(* IEC 61131-3 sources: test/Class/LseEasy, 1 file *)

(* ---- LseEasy.st ---- *)
#include "..\..\Source\Common\hmi_nuc.h"

(*!
<Class
	Name               = "LseEasy"
	Revision           = "1.32"
	RealtimeTask       = "false"
	CyclicTask         = "false"
	BackgroundTask     = "true"
	DefBackground      = "always"
	Sigmatek           = "true"
	OSInterface        = "false"
	HighPriority       = "false"
	Automatic          = "false"
	UpdateMode         = "Prescan"
	SharedCommandTable = "true"
	Objectsize         = "(474,120)"
	Comment            = "Class is used to operate LSE-Easy Visualization&#13;&#10;LSE-CompilerVersion: 60">
	<Channels>
		<Server Name="AccessLevel" Visualized="true" Initialize="false" WriteProtected="false" Retentive="false" Comment="server is used to disable/enable access to several inputs and buttons&#13;&#10;virtual method HmiAccess() is responsible for algorithm."/>
		<Server Name="ActHumidity" Visualized="true" Initialize="false" WriteProtected="true" Retentive="false" Comment="actual humidity"/>
		<Server Name="ActLanguage" Visualized="true" Initialize="true" DefValue="0" WriteProtected="false" Retentive="SRam" Comment="Server is used to select language&#13;&#10;use index or accurate language designator to switch over"/>
		<Server Name="ActScreen" Visualized="true" Initialize="false" WriteProtected="false" Retentive="false" Comment="server is used to show number of actual screen on hmi&#13;&#10;call write-method with accurate screennumber given by lse to force hmi to view new screen&#13;&#10;call writemethode with -2 to get screenshot from hmi (C:\hmi35.bmp)"/>
		<Server Name="ActTemperature" Visualized="true" Initialize="false" WriteProtected="true" Retentive="false" Comment="actual temperature"/>
		<Server Name="BacklightDim" Visualized="true" Initialize="false" WriteProtected="false" Retentive="false" Comment="server is used to dim backlight of hmi&#13;&#10;call writemethode with any value from 0 to 100 to dim backlight&#13;&#10;0 .... next to dark&#13;&#10;100 .. bright"/>
		<Server Name="BacklightOnOff" Visualized="false" Initialize="false" WriteProtected="false" Retentive="false" Comment="server is used to turn on/off backlight of hmi&#13;&#10;call writemethode with 0 to turn off backlight&#13;&#10;on the oter hand call writemethode with 1 to turn on backlight"/>
		<Server Name="ClassSvr" Visualized="false" Initialize="false" WriteProtected="true" Retentive="false"/>
		<Server Name="ErrorSvr" Visualized="true" Initialize="false" WriteProtected="true" Retentive="false"/>
		<Server Name="HmiHwVersion" Visualized="true" Initialize="false" WriteProtected="true" Retentive="false" Comment="is used to view hardwareversion of hmi"/>
		<Server Name="HmiOnline" Visualized="true" Initialize="false" WriteProtected="true" Retentive="false" Comment="0 ... hmi is offline&#13;&#10;1 ... hmi is online"/>
		<Server Name="HmiSwVersion" Visualized="true" Initialize="false" WriteProtected="true" Retentive="false" Comment="is used to view softwareversion (firmware) of hmi"/>
		<Server Name="LastUsage" Visualized="false" Initialize="false" WriteProtected="true" Retentive="false" Comment="server is used to display timestamp (ops.tabsolute) of last usage of hmi"/>
		<Server Name="ListVal0" Visualized="true" Initialize="false" WriteProtected="false" Retentive="false" Comment="server is used to display arbitrary scrolllist on display&#13;&#10;actual selection in list will be shown on server"/>
		<Server Name="ListVal1" Visualized="true" Initialize="false" WriteProtected="false" Retentive="false"/>
		<Server Name="LseProjectRevision" Visualized="true" Initialize="false" WriteProtected="true" Retentive="false"/>
		<Server Name="PixMap" Visualized="true" Initialize="false" WriteProtected="false" Retentive="false"/>
		<Server Name="StateSvr" Visualized="true" Initialize="false" WriteProtected="false" Retentive="false" Comment="actual state of program"/>
		<Server Name="TrendVal0" Visualized="true" Initialize="false" WriteProtected="false" Retentive="false" Comment="server is used to display trend0 on hmi&#13;&#10;call writemethod with any value from 0 to 255 to add value"/>
		<Server Name="TrendVal1" Visualized="true" Initialize="false" WriteProtected="false" Retentive="false" Comment="server is used to display trend1 on hmi&#13;&#10;call writemethod with any value from 0 to 255 to add value"/>
		<Client Name="AutoFirmwareUpdate" Required="true" Internal="false" DefValue="0" Comment="Client is used to ensure automatic update of firmware and bootloader at hmi after poweron of connected plc.&#13;&#10;Set client to 1 or 2 to enable automatic update otherwirse, when client is set to 0, automatic update is disabled.&#13;&#10;NOTE: &#13;&#10;If client is set to 1, updatefiles will be deleted after update of hmi. &#13;&#10;When client is set to 2, updatefiles will NOT be deleted after automatic update. In that case user has to disconnect device otherwise update will be performed each time after poweron.&#13;&#10;User has to place updatefiles at correct device (eg.: C:\, E:\, ...}. When updatefiles should be deleted after success make sure that device and updatefiles are not writeprotected.&#13;&#10;Use virtual methods GetUpdatePath(), GetFirmwareUpdate() and GetBootLoaderUpdate() to customize device, directory and name of updatefiles."/>
		<Client Name="BackLightOff" Required="true" Internal="false" DefValue="300000" Comment="client is used to set duration till backlight will be turned off when display is not in use&#13;&#10;timebase is milliseconds&#13;&#10;0 ... backlight is always on"/>
		<Client Name="ComPort" Required="true" Internal="false" Comment="client is used to communicate with hmi&#13;&#10;eg: connect instance of class HmiComPortCan to communicate vie canbus"/>
		<Client Name="File" Required="true" Internal="true"/>
		<Client Name="HmiChkBitList" Required="true" Internal="true"/>
		<Client Name="HmiColorMap" Required="true" Internal="true"/>
		<Client Name="HmiFont35" Required="true" Internal="true"/>
		<Client Name="HmiFontList" Required="true" Internal="true"/>
		<Client Name="HmiFontShemeList" Required="true" Internal="true"/>
		<Client Name="HmiFunctionList" Required="true" Internal="true"/>
		<Client Name="HmiFunctionList35" Required="true" Internal="true"/>
		<Client Name="HmiImage35" Required="true" Internal="true"/>
		<Client Name="HmiImageList" Required="true" Internal="true"/>
		<Client Name="HmiImageShemeList" Required="true" Internal="true"/>
		<Client Name="HmiMapFile" Required="true" Internal="true"/>
		<Client Name="HmiProject35" Required="true" Internal="true"/>
		<Client Name="HmiProjectList" Required="true" Internal="true"/>
		<Client Name="HmiScreen" Required="true" Internal="true"/>
		<Client Name="HmiSetUpList" Required="true" Internal="true"/>
		<Client Name="HmiSetupList35" Required="true" Internal="true"/>
		<Client Name="HmiShemeList35" Required="true" Internal="true"/>
		<Client Name="HmiStateBit35" Required="true" Internal="true"/>
		<Client Name="HmiT9Config" Required="true" Internal="true"/>
		<Client Name="HmiTextList" Required="true" Internal="true"/>
		<Client Name="HmiTextList35" Required="true" Internal="true"/>
		<Client Name="HmiTextShemeList" Required="true" Internal="true"/>
		<Client Name="HmiUtils" Required="true" Internal="true"/>
		<Client Name="HmiVarList" Required="true" Internal="true"/>
		<Client Name="HmiVarList35" Required="true" Internal="true"/>
		<Client Name="OverloadLight" Required="true" Internal="false" DefValue="-1" Comment="client is used to ensure overload&#13;&#10;if client is set to equal or bigger 0 all occurences of &quot;XX&quot; in variablename done with LSE will be xchanged with adequateness number of client"/>
		<Client Name="ProjectPath" Required="true" Internal="false" DefValue="0" Comment="selector for different projectpath&#13;&#10;0: C:\MPC\&#13;&#10;&gt;0: C:\Easy[Value]\ (eg.: C:\Easy123\)&#13;&#10;-1: C:\[ObjextName]\ (eg.: C:\LSEEASY1\)&#13;&#10;"/>
		<Client Name="StringLib" Required="true" Internal="true"/>
		<Client Name="TempInterval" Required="true" Internal="false" DefValue="1000" Comment="client is used to define interval of retrieving act.temperature from hmi&#13;&#10;timebase is milliseconds&#13;&#10;0 ... do not update act.temperature"/>
	</Channels>
	<Dependencies>
		<Files>
			<File Path=".\Source\Common\hmi_nuc.h" Include="true"/>
			<File Path=".\Class\LseEasy\MiniSrcData.h" Include="false"/>
			<File Path=".\Class\LseEasy\Create.h" Include="false"/>
			<File Path=".\Class\LseEasy\CreateScreen.c"/>
			<File Path=".\Class\LseEasy\CreateUtils.c"/>
		</Files>
	</Dependencies>
	<RevDoku>
		<Owner Company="sigmatek" Author="kolott"/>
		<Dokumentation Revision="1.32" Date="2021-02-26" Author="kolott" Company="sigmatek" Description="Method LseEasy::ListSetup() by parameter &apos;bottom_up&apos; expanded&#13;&#10;8D-1972: Extended size of textpuffer"/>
		<Dokumentation Revision="1.31" Date="2020-04-28" Author="kolott" Company="sigmatek" Description="New method GetLseProjectName() added&#13;&#10;DEVVIS-40, sa57116: New method T9KeyboardConfig() added"/>
		<Dokumentation Revision="1.30" Date="2019-01-24" Author="kolott" Company="sigmatek" Description="Support of HZS-251-1 and HZS352-1 incl. Humidity"/>
		<Dokumentation Revision="1.29" Date="2019-01-09" Author="kolott" Company="sigmatek" Description="Virtual method HmiOverloadLight() added to ensure userspecific change of Objectname"/>
		<Dokumentation Revision="1.28" Date="2018-10-18" Author="kolott" Company="sigmatek" Description="sa42417: more than 6 different projectpath implemented in virtual method LseEasy::GetPrjPath()"/>
		<Dokumentation Revision="1.27" Date="2018-08-27" Author="kolott" Company="sigmatek" Description="Problem &quot;Out Of Memory&quot; will end in Error &quot;Can&apos;t load LSE-Project&quot;&#13;&#10;Variable Limits at Variables will work. Overwrite Method LseEasy::VariableLimitsInUse() to enable feature"/>
		<Dokumentation Revision="1.26" Date="2018-05-24" Author="kolott" Company="sigmatek" Description="sa41119, DEVSW502: Send individual StandardFonts given by LSE to HMI as well. Fonts are used in Standard Keypads"/>
		<Dokumentation Revision="1.25" Date="2018-04-18" Author="kolott" Company="sigmatek" Description="sa40364: userspecific xchange of images done by LSE.&#13;&#10;DEVSW440: Server ActTemperature is set to 16#80000010 when HMI is offline and TemperatureValue is needed"/>
		<Dokumentation Revision="1.24" Date="2018-01-17" Author="kolott" Company="sigmatek" Description="TextList done wilt LSE will be accessible by user during runtime&#13;&#10;new virtual method HmiProjectBegin(), AddVariableByName() and AddStateBitByName() added"/>
		<Dokumentation Revision="1.23" Date="2016-09-07" Author="kolott" Company="sigmatek" Description="sa35391: new method GetLseProjectNotice() and Server LseProjectRevision added&#13;&#10;sa35411: correction in entire bytesizecomputation of HMI-project-data"/>
		<Dokumentation Revision="1.22" Date="2016-07-08" Author="kolott" Company="sigmatek" Description="new Client AutoFirmwareUpdate added to enable automatic update of firmware and bootloader at hmi after poweron"/>
		<Dokumentation Revision="1.21" Date="2016-06-22" Author="kolott" Company="sigmatek" Description="Functionality to Update BootLoader in HMI added"/>
		<Dokumentation Revision="1.20" Date="2016-05-03" Author="kolott" Company="sigmatek" Description="Betterment in rounding result at method Calc().&#13;&#10;Set and resetvalue at button will work. Firmwareversion 1.35 or higher is necessary at HMI.&#13;&#10;sa26785: compilerversion 60, property preceding zero implemented&#13;&#10;Methode UpdateString35() is done virtual"/>
		<Dokumentation Revision="1.19" Date="2016-04-23" Author="kolott" Company="sigmatek" Description="sa34276: new methode Recalculate() added to ensure recalculation from binary to physical values"/>
		<Dokumentation Revision="1.18" Date="2016-03-12" Author="kolott" Company="sigmatek" Description="functionality to display pixmap (barcode, qr code,...) on hmi added. use method SendPixMap() to view data&#13;&#10;correction of server ActLanguage when actual selection doesn&apos;t fit to loaded project (sa33823)"/>
		<Dokumentation Revision="1.17" Date="2016-02-04" Author="kolott" Company="sigmatek" Description="new virtual method IsProjectUpLoadNecessary() to customize project-upload added"/>
		<Dokumentation Revision="1.16" Date="2015-11-30" Author="kolott" Company="sigmatek" Description="new Server &quot;ListVal1&quot; to ensure use of second scrolllist on HMI"/>
		<Dokumentation Revision="1.15" Date="2015-03-17" Author="kolott" Company="sigmatek" Description="method UpdateValue35() is done &quot;virtual&quot;"/>
		<Dokumentation Revision="1.14" Date="2014-11-26" Author="kolott" Company="sigmatek" Description="new method HmiVariableExtention() used to ensure userextended modifications done in firmware of hmi&#13;&#10;view Passwordcharacter at String will work"/>
		<Dokumentation Revision="1.13" Date="2014-10-15" Author="kolott" Company="sigmatek" Description="Ability to customise HmiProject added (HmiProjectCreate(), CreateAddText(), CreateAddImage(), ListSetup(), ListCmd(), ListAddItem())"/>
		<Dokumentation Revision="1.12" Date="2014-08-13" Author="kolott" Company="sigmatek" Description="Server &quot;ListVal0&quot; is added to ensure scrollist on HMI&#13;&#10;Function &quot;UserCall&quot; added&#13;&#10;Retry added at filetransfer to HMI"/>
		<Dokumentation Revision="1.11" Date="2014-08-07" Author="kolott" Company="sigmatek" Description="Server of type ENUM will work as well"/>
		<Dokumentation Revision="1.10" Date="2014-06-02" Author="kolott" Company="sigmatek" Description="Method &quot;UpdateTemperature35&quot; is virtual to ensure correction of actual HMI-Temperature&#13;&#10;Correction: Display of Unicode-String always started with character &apos;?&apos;"/>
		<Dokumentation Revision="1.9" Date="2014-04-28" Author="kolott" Company="sigmatek" Description="call of function &quot;Function Block&quot; activated&#13;&#10;view of Circle + Pie added"/>
		<Dokumentation Revision="1.8" Date="2014-04-14" Author="kolott" Company="sigmatek" Description="betterment in Offline-Mode when HMI (display) is not connected&#13;&#10;new virtual method GetFirmwareUpdate() to customize drive and name of firmwareupdatefile&#13;&#10;reduce of memoryrequirement in plc"/>
		<Dokumentation Revision="1.7" Date="2014-03-26" Author="kolott" Company="sigmatek" Description="attribute bold at text will work as well when firmwareversion &gt;= 1.24 is in use&#13;&#10;DownloadOnTheFly will work with accurate LSE-Version"/>
		<Dokumentation Revision="1.6" Date="2014-03-06" Author="kolott" Company="sigmatek" Description="accesslevel and chkbits will work&#13;&#10;new Server AccessLevel&#13;&#10;EasyMap.xml instead of EasyMap.txt will be generated"/>
		<Dokumentation Revision="1.5" Date="2014-02-27" Author="kolott" Company="sigmatek" Description="more than one hmi with different lse-projects are possible"/>
		<Dokumentation Revision="1.4" Date="2014-02-27" Author="kolott" Company="sigmatek" Description="variable limits at bar (hmi-firmware 1.22)&#13;&#10;slider (bar + writeprotect = false) (hmi-firmware 1.22)&#13;&#10;zoomable imagescheme"/>
		<Dokumentation Revision="1.3" Date="2014-02-13" Author="kolott" Company="sigmatek" Description="Server ErrorSvr to view errordetails added"/>
		<Dokumentation Revision="1.2" Date="2014-02-12" Author="kolott" Company="sigmatek" Description="server LastUsage added"/>
		<Dokumentation Revision="1.1" Date="2014-01-16" Author="kolott" Company="sigmatek" Description="Trend added"/>
		<Dokumentation Revision="1.0" Date="2013-12-19" Author="kolott" Company="sigmatek" Description="release"/>
	</RevDoku>
	<Network Name="LseEasy">
		<!-- List of Components in this network -->
		<Components>
			<Object
				Name       = "File"
				Class      = "HmiFile"
				Position   = "(90,720)"
				Visualized = "false">
				<Channels>
					<Server Name="ClassSvr"/>
					<Client Name="OpSysFile"/>
					<Client Name="StdLib"/>
				</Channels>
			</Object>
			<Object
				Name       = "HmiChkBitList"
				Class      = "HmiChkBitList"
				Position   = "(1050,330)"
				Visualized = "false">
				<Channels>
					<Server Name="ClassSvr"/>
					<Client Name="File"/>
					<Client Name="StringLib"/>
					<Client Name="VarList"/>
				</Channels>
			</Object>
			<Object
				Name       = "HmiColorMap"
				Class      = "HmiColorMap"
				Position   = "(540,390)"
				Visualized = "false">
				<Channels>
					<Server Name="ClassSvr"/>
					<Client Name="File"/>
				</Channels>
			</Object>
			<Object
				Name       = "HmiFont35"
				Class      = "HmiFont35"
				Position   = "(1530,1620)"
				Visualized = "false">
				<Channels>
					<Server Name="ByteSize"/>
					<Server Name="ClassSvr"/>
					<Client Name="StdLib"/>
				</Channels>
			</Object>
			<Object
				Name       = "HmiFontList"
				Class      = "HmiFontList"
				Position   = "(540,1050)"
				Visualized = "false">
				<Channels>
					<Server Name="ClassSvr"/>
					<Client Name="File"/>
					<Client Name="StringLib"/>
				</Channels>
			</Object>
			<Object
				Name       = "HmiFontShemeList"
				Class      = "HmiShemeList"
				Position   = "(540,540)"
				Visualized = "false">
				<Channels>
					<Server Name="ClassSvr"/>
					<Client Name="File"/>
				</Channels>
			</Object>
			<Object
				Name       = "HmiFunctionList"
				Class      = "HmiFunctionList"
				Position   = "(540,900)"
				Visualized = "false">
				<Channels>
					<Server Name="ClassSvr"/>
					<Client Name="File"/>
				</Channels>
			</Object>
			<Object
				Name       = "HmiFunctionList35"
				Class      = "HmiFunctionList35"
				Position   = "(1050,1830)"
				Visualized = "false">
				<Channels>
					<Server Name="ByteSize"/>
					<Server Name="ClassSvr"/>
					<Client Name="HmiVarList"/>
				</Channels>
			</Object>
			<Object
				Name       = "HmiImage35"
				Class      = "HmiImage35"
				Position   = "(1530,1830)"
				Visualized = "false">
				<Channels>
					<Server Name="ByteSize"/>
					<Server Name="ClassSvr"/>
					<Client Name="StdLib"/>
				</Channels>
			</Object>
			<Object
				Name       = "HmiImageList"
				Class      = "HmiImageList"
				Position   = "(540,690)"
				Visualized = "false">
				<Channels>
					<Server Name="ClassSvr"/>
					<Client Name="File"/>
					<Client Name="StringLib"/>
				</Channels>
			</Object>
			<Object
				Name       = "HmiImageShemeList"
				Class      = "HmiShemeList"
				Position   = "(1530,660)"
				Visualized = "false">
				<Channels>
					<Server Name="ClassSvr"/>
					<Client Name="File"/>
				</Channels>
			</Object>
			<Object
				Name       = "HmiMapFile"
				Class      = "HmiMapFile"
				Position   = "(1530,1050)"
				Visualized = "false">
				<Channels>
					<Server Name="ClassSvr"/>
					<Client Name="File"/>
					<Client Name="StateBit"/>
					<Client Name="StringLib"/>
					<Client Name="VarList"/>
				</Channels>
			</Object>
			<Object
				Name       = "HmiProject35"
				Class      = "HmiProject35"
				Position   = "(90,1560)"
				Visualized = "false">
				<Channels>
					<Server Name="ClassSvr"/>
					<Server Name="TotalByteSize"/>
					<Server Name="TotalFileNo"/>
					<Client Name="StdLib"/>
				</Channels>
			</Object>
			<Object
				Name       = "HmiProjectList"
				Class      = "HmiProjectList"
				Position   = "(540,180)"
				Visualized = "false">
				<Channels>
					<Server Name="ClassSvr"/>
					<Client Name="File"/>
					<Client Name="StringLib"/>
				</Channels>
			</Object>
			<Object
				Name       = "HmiScreen"
				Class      = "HmiScreen"
				Position   = "(1530,180)"
				Visualized = "false">
				<Channels>
					<Server Name="ClassSvr"/>
					<Client Name="File"/>
				</Channels>
			</Object>
			<Object
				Name       = "HmiSetUpList"
				Class      = "HmiSetUpList"
				Position   = "(1050,180)"
				Visualized = "false">
				<Channels>
					<Server Name="ClassSvr"/>
					<Client Name="File"/>
				</Channels>
			</Object>
			<Object
				Name       = "HmiSetupList35"
				Class      = "HmiSetupList35"
				Position   = "(90,1830)"
				Visualized = "false">
				<Channels>
					<Server Name="ByteSize"/>
					<Server Name="ClassSvr"/>
				</Channels>
			</Object>
			<Object
				Name       = "HmiShemeList35"
				Class      = "HmiShemeList35"
				Position   = "(540,1830)"
				Visualized = "false">
				<Channels>
					<Server Name="ByteSize"/>
					<Server Name="ClassSvr"/>
				</Channels>
			</Object>
			<Object
				Name       = "HmiStateBit35"
				Class      = "HmiStateBit35"
				Position   = "(1050,1050)"
				Visualized = "false">
				<Channels>
					<Server Name="ClassSvr"/>
					<Client Name="ChkBit"/>
					<Client Name="ComPort"/>
					<Client Name="StringLib"/>
					<Client Name="VarList"/>
				</Channels>
			</Object>
			<Object
				Name       = "HmiT9Config"
				Class      = "HmiT9Config35"
				Position   = "(540,1410)"
				Visualized = "false">
				<Channels>
					<Server Name="ByteSize"/>
					<Server Name="ClassSvr"/>
				</Channels>
			</Object>
			<Object
				Name       = "HmiTextList"
				Class      = "HmiTextList"
				Position   = "(1530,330)"
				Visualized = "false">
				<Channels>
					<Server Name="ClassSvr"/>
					<Client Name="File"/>
					<Client Name="HmiTextList35"/>
					<Client Name="HmiVarList"/>
					<Client Name="StringLib"/>
				</Channels>
			</Object>
			<Object
				Name       = "HmiTextList35"
				Class      = "HmiTextList35"
				Position   = "(1050,1620)"
				Visualized = "false">
				<Channels>
					<Server Name="ByteSize"/>
					<Server Name="ClassSvr"/>
				</Channels>
			</Object>
			<Object
				Name       = "HmiTextShemeList"
				Class      = "HmiShemeList"
				Position   = "(1530,810)"
				Visualized = "false">
				<Channels>
					<Server Name="ClassSvr"/>
					<Client Name="File"/>
				</Channels>
			</Object>
			<Object
				Name       = "HmiUtils"
				Class      = "HmiUtils"
				Position   = "(90,570)"
				Visualized = "false">
				<Channels>
					<Server Name="ClassSvr"/>
				</Channels>
			</Object>
			<Object
				Name       = "HmiVarList"
				Class      = "HmiVarList"
				Position   = "(1050,630)"
				Visualized = "false">
				<Channels>
					<Server Name="ClassSvr"/>
					<Client Name="ComPort"/>
					<Client Name="File"/>
					<Client Name="HmiVarList35"/>
					<Client Name="StringLib"/>
					<Client Name="TextList"/>
				</Channels>
			</Object>
			<Object
				Name       = "HmiVarList35"
				Class      = "HmiVarList35"
				Position   = "(540,1620)"
				Visualized = "false">
				<Channels>
					<Server Name="ByteSize"/>
					<Server Name="ClassSvr"/>
				</Channels>
			</Object>
			<Object
				Name       = "StringLib"
				Class      = "HmiStrLib"
				Position   = "(90,930)"
				Visualized = "false">
				<Channels>
					<Server Name="ClassSvr"/>
					<Client Name="StdLib"/>
				</Channels>
			</Object>
		</Components>
		<Comments>
		</Comments>
		<!-- List of Connections in this network -->
		<Connections>
			<Connection Source="this.HmiImageList" Destination="HmiImageList.ClassSvr"/>
			<Connection Source="this.File" Destination="File.ClassSvr"/>
			<Connection Source="this.HmiVarList" Destination="HmiVarList.ClassSvr"/>
			<Connection Source="HmiProjectList.File" Destination="File.ClassSvr" Vertices="(540,270),(450,270),(450,810),(390,810),"/>
			<Connection Source="this.HmiFunctionList" Destination="HmiFunctionList.ClassSvr"/>
			<Connection Source="HmiColorMap.File" Destination="File.ClassSvr" Vertices="(540,480),(450,480),(450,810),(390,810),"/>
			<Connection Source="this.StringLib" Destination="StringLib.ClassSvr"/>
			<Connection Source="this.HmiScreen" Destination="HmiScreen.ClassSvr"/>
			<Connection Source="HmiFontShemeList.File" Destination="File.ClassSvr" Vertices="(540,630),(450,630),(450,810),(390,810),"/>
			<Connection Source="this.HmiTextList" Destination="HmiTextList.ClassSvr"/>
			<Connection Source="HmiImageList.File" Destination="File.ClassSvr" Vertices="(540,780),(450,780),(450,810),(390,810),"/>
			<Connection Source="HmiFunctionList.File" Destination="File.ClassSvr" Vertices="(540,990),(450,990),(450,810),(390,810),"/>
			<Connection Source="this.HmiImageShemeList" Destination="HmiImageShemeList.ClassSvr"/>
			<Connection Source="this.HmiTextShemeList" Destination="HmiTextShemeList.ClassSvr"/>
			<Connection Source="HmiFontList.File" Destination="File.ClassSvr" Vertices="(540,1140),(450,1140),(450,810),(390,810),"/>
			<Connection Source="HmiSetUpList.File" Destination="File.ClassSvr" Vertices="(1050,270),(930,270),(930,120),(450,120),(450,810),(390,810),"/>
			<Connection Source="this.HmiFontShemeList" Destination="HmiFontShemeList.ClassSvr"/>
			<Connection Source="HmiScreen.File" Destination="File.ClassSvr" Vertices="(1530,270),(1470,270),(1470,120),(450,120),(450,810),(390,810),"/>
			<Connection Source="this.HmiFontList" Destination="HmiFontList.ClassSvr"/>
			<Connection Source="HmiTextList.File" Destination="File.ClassSvr" Vertices="(1530,420),(1470,420),(1470,120),(450,120),(450,810),(390,810),"/>
			<Connection Source="HmiImageShemeList.File" Destination="File.ClassSvr" Vertices="(1530,750),(1470,750),(1470,120),(450,120),(450,810),(390,810),"/>
			<Connection Source="this.HmiColorMap" Destination="HmiColorMap.ClassSvr"/>
			<Connection Source="HmiTextShemeList.File" Destination="File.ClassSvr" Vertices="(1530,900),(1470,900),(1470,120),(450,120),(450,810),(390,810),"/>
			<Connection Source="this.HmiProjectList" Destination="HmiProjectList.ClassSvr"/>
			<Connection Source="HmiVarList.File" Destination="File.ClassSvr" Vertices="(1050,720),(930,720),(930,120),(450,120),(450,810),(390,810),"/>
			<Connection Source="HmiTextList.StringLib" Destination="StringLib.ClassSvr" Vertices="(1530,480),(1440,480),(1440,150),(480,150),(480,1020),(390,1020),"/>
			<Connection Source="HmiVarList.TextList" Destination="HmiTextList.ClassSvr" Vertices="(1050,840),(1830,420),"/>
			<Connection Source="this.HmiProject35" Destination="HmiProject35.ClassSvr"/>
			<Connection Source="this.HmiVarList35" Destination="HmiVarList35.ClassSvr"/>
			<Connection Source="HmiVarList.HmiVarList35" Destination="HmiVarList35.ClassSvr" Vertices="(1050,900),(930,900),(930,1710),(840,1710),"/>
			<Connection Source="this.HmiFont35" Destination="HmiFont35.ClassSvr"/>
			<Connection Source="HmiTextList.HmiVarList" Destination="HmiVarList.ClassSvr" Vertices="(1530,540),(1380,540),(1380,720),(1350,720),"/>
			<Connection Source="this.HmiImage35" Destination="HmiImage35.ClassSvr"/>
			<Connection Source="this.HmiSetUpList" Destination="HmiSetUpList.ClassSvr"/>
			<Connection Source="HmiProjectList.StringLib" Destination="StringLib.ClassSvr" Vertices="(540,330),(480,330),(480,1020),(390,1020),"/>
			<Connection Source="this.HmiFunctionList35" Destination="HmiFunctionList35.ClassSvr"/>
			<Connection Source="HmiFunctionList35.HmiVarList" Destination="HmiVarList.ClassSvr" Vertices="(1050,1920),(990,1920),(990,1470),(1380,1470),(1380,720),(1350,720),"/>
			<Connection Source="this.HmiShemeList35" Destination="HmiShemeList35.ClassSvr"/>
			<Connection Source="HmiVarList.ComPort" Destination="this.ComPort" Vertices="(1050,960),(38,210),"/>
			<Connection Source="this.HmiSetupList35" Destination="HmiSetupList35.ClassSvr"/>
			<Connection Source="HmiImageList.StringLib" Destination="StringLib.ClassSvr" Vertices="(540,840),(480,840),(480,1020),(390,1020),"/>
			<Connection Source="HmiFontList.StringLib" Destination="StringLib.ClassSvr" Vertices="(540,1200),(480,1200),(480,1020),(390,1020),"/>
			<Connection Source="HmiVarList.StringLib" Destination="StringLib.ClassSvr" Vertices="(1050,780),(960,780),(960,150),(480,150),(480,1020),(390,1020),"/>
			<Connection Source="this.HmiUtils" Destination="HmiUtils.ClassSvr"/>
			<Connection Source="this.HmiTextList35" Destination="HmiTextList35.ClassSvr"/>
			<Connection Source="HmiTextList.HmiTextList35" Destination="HmiTextList35.ClassSvr" Vertices="(1530,600),(1410,600),(1410,1710),(1350,1710),"/>
			<Connection Source="this.HmiChkBitList" Destination="HmiChkBitList.ClassSvr"/>
			<Connection Source="HmiChkBitList.File" Destination="File.ClassSvr" Vertices="(1050,420),(930,420),(930,120),(450,120),(450,810),(390,810),"/>
			<Connection Source="HmiChkBitList.VarList" Destination="HmiVarList.ClassSvr" Vertices="(1050,480),(990,480),(990,600),(1380,600),(1380,720),(1350,720),"/>
			<Connection Source="this.HmiStateBit35" Destination="HmiStateBit35.ClassSvr"/>
			<Connection Source="HmiStateBit35.ChkBit" Destination="HmiChkBitList.ClassSvr" Vertices="(1050,1140),(1350,420),"/>
			<Connection Source="HmiStateBit35.ComPort" Destination="this.ComPort" Vertices="(1050,1200),(38,210),"/>
			<Connection Source="HmiStateBit35.VarList" Destination="HmiVarList.ClassSvr" Vertices="(1050,1260),(990,1260),(990,1020),(1380,1020),(1380,720),(1350,720),"/>
			<Connection Source="this.HmiMapFile" Destination="HmiMapFile.ClassSvr"/>
			<Connection Source="HmiMapFile.File" Destination="File.ClassSvr" Vertices="(1530,1140),(1470,1140),(1470,120),(450,120),(450,810),(390,810),"/>
			<Connection Source="HmiMapFile.VarList" Destination="HmiVarList.ClassSvr" Vertices="(1530,1200),(1380,1200),(1380,720),(1350,720),"/>
			<Connection Source="HmiMapFile.StateBit" Destination="HmiStateBit35.ClassSvr" Vertices="(1530,1260),(1350,1140),"/>
			<Connection Source="HmiMapFile.StringLib" Destination="StringLib.ClassSvr" Vertices="(1530,1320),(1440,1320),(1440,150),(480,150),(480,1020),(390,1020),"/>
			<Connection Source="HmiStateBit35.StringLib" Destination="StringLib.ClassSvr" Vertices="(1050,1320),(960,1320),(960,150),(480,150),(480,1020),(390,1020),"/>
			<Connection Source="HmiChkBitList.StringLib" Destination="StringLib.ClassSvr" Vertices="(1050,540),(960,540),(960,150),(480,150),(480,1020),(390,1020),"/>
			<Connection Source="this.HmiT9Config" Destination="HmiT9Config.ClassSvr"/>
		</Connections>
		<!-- Headerfiles -->
		<Options>
		</Options>
	</Network>
</Class>
*)
LseEasy : CLASS
	TYPE
	  TErrorSvr :  //! <Type Public="true" Name="TErrorSvr"/>
	  (
	    ErrNone,
	    ErrCreateHmiProject,
	    ErrLseCompilerVersion,
	    ErrLoadLseProject,
	    ErrSizeLseProject,
	    ErrUploadHmiProject,
	    ErrHmiCommunication
	  )$UDINT;
	  TStateSvr :  //! <Type Public="true" Name="TStateSvr"/>
	  (
	    TStart,
	    TUpLoad,
	    TRun,
	    TError,
	    TFirmwareUpdate,
	    TSleep,
	    TChkCrc,
	    TGetScreenShot,
	    TReboot,
	    TBootLoaderUpdate,
	    TCheckUpdateBootloader,
	    TCheckUpdateFirmware
	  )$UDINT;
	END_TYPE
  //Servers:
	ClassSvr 	: SvrChCmd_DINT;
	StateSvr 	: SvrCh_TStateSvr_PTofCls_LseEasy;
	ErrorSvr 	: SvrCh_TErrorSvr_PTofCls_LseEasy;
	HmiOnline 	: SvrCh_DINT;
	ActTemperature 	: SvrCh_DINT;
	ActLanguage 	: SvrCh_UDINT;
	ActScreen 	: SvrCh_DINT;
	BacklightOnOff 	: SvrCh_DINT;
	BacklightDim 	: SvrCh_DINT;
	TrendVal0 	: SvrCh_DINT;
	TrendVal1 	: SvrCh_DINT;
	LastUsage 	: SvrCh_UDINT;
	HmiSwVersion 	: SvrCh_UDINT;
	HmiHwVersion 	: SvrCh_UDINT;
	AccessLevel 	: SvrCh_UDINT;
	ListVal0 	: SvrCh_DINT;
	ListVal1 	: SvrCh_DINT;
	PixMap 	: SvrCh_DINT;
	LseProjectRevision 	: SvrCh_HDINT;
	ActHumidity 	: SvrCh_DINT;
  //Clients:
	ComPort 	: CltChCmd_HmiComPort;
	HmiImageList 	: CltChCmd_HmiImageList;
	HmiFunctionList 	: CltChCmd_HmiFunctionList;
	HmiScreen 	: CltChCmd_HmiScreen;
	HmiFontList 	: CltChCmd_HmiFontList;
	HmiVarList 	: CltChCmd_HmiVarList;
	HmiColorMap 	: CltChCmd_HmiColorMap;
	HmiProjectList 	: CltChCmd_HmiProjectList;
	HmiProject35 	: CltChCmd_HmiProject35;
	HmiTextList 	: CltChCmd_HmiTextList;
	HmiVarList35 	: CltChCmd_HmiVarList35;
	HmiFont35 	: CltChCmd_HmiFont35;
	HmiImage35 	: CltChCmd_HmiImage35;
	HmiSetUpList 	: CltChCmd_HmiSetUpList;
	HmiFunctionList35 	: CltChCmd_HmiFunctionList35;
	HmiShemeList35 	: CltChCmd_HmiShemeList35;
	HmiFontShemeList 	: CltChCmd_HmiShemeList;
	ProjectPath 	: CltCh_DINT;
	TempInterval 	: CltCh_UDINT;
	BackLightOff 	: CltCh_UDINT;
	HmiTextShemeList 	: CltChCmd_HmiShemeList;
	HmiImageShemeList 	: CltChCmd_HmiShemeList;
	HmiSetupList35 	: CltChCmd_HmiSetupList35;
	StringLib 	: CltChCmd_HmiStrLib;
	File 	: CltChCmd_HmiFile;
	HmiUtils 	: CltChCmd_HmiUtils;
	OverloadLight 	: CltCh_DINT;
	HmiTextList35 	: CltChCmd_HmiTextList35;
	HmiChkBitList 	: CltChCmd_HmiChkBitList;
	HmiStateBit35 	: CltChCmd_HmiStateBit35;
	HmiMapFile 	: CltChCmd_HmiMapFile;
	AutoFirmwareUpdate 	: CltCh_DINT;
	HmiT9Config 	: CltChCmd_HmiT9Config35;
  //Variables:
		ProjectBox 	: ^void;
		AliveTix35Cntr 	: UDINT;
		AliveTix35CntrOld 	: UDINT;
		AliveTix35 	: UDINT;
		AliveTix 	: UDINT;
		HmiPrjCrc 	: UDINT;
		Hmi35PrjCrc 	: UDINT;
		RefreshTix 	: UDINT;
		StateNext 	: TStateSvr;
		TrendVal0Lid 	: UDINT;
		TrendVal1Lid 	: UDINT;
		TryToRestart 	: BOOL;
		CallScreen 	: DINT;
		NeedUpdateAll 	: UDINT;
		CantGetCrc 	: UDINT;
		SleepStart 	: UDINT;
		SleepDuration 	: UDINT;
		BacklightDimLid 	: UDINT;
		HmiSwVersionLid 	: UDINT;
		HmiHwVersionLid 	: UDINT;
		ListVal0Lid 	: UDINT;
		ListVal1Lid 	: UDINT;
		CreateAdd 	: BOOL;
		PixMapLid 	: UDINT;
		TmpData : ARRAY [0..3000] OF USINT;

		UpdateFileDPNE : ARRAY [0..255] OF CHAR;

		AutoFwUpdateDisabled 	: BOOL;
		LseProjectPath : ARRAY [0..32] OF CHAR;

  //Functions:

	FUNCTION LseEasy
		VAR_OUTPUT
			ret_code 	: ConfStates;
		END_VAR;

	FUNCTION VIRTUAL GLOBAL Init;

	FUNCTION VIRTUAL GLOBAL Background
		VAR_INPUT
			EAX 	: UDINT;
		END_VAR
		VAR_OUTPUT
			state (EAX) 	: UDINT;
		END_VAR;

	FUNCTION LoadFile
		VAR_OUTPUT
			retcode 	: BOOL;
		END_VAR;
				//! <Function Comment="method is used to serve projectpath" Name="GetPrjPath"/>
	FUNCTION VIRTUAL GLOBAL GetPrjPath
		VAR_OUTPUT
			retcode 	: ^LASCII;
		END_VAR;

	FUNCTION MakePrjFileName
		VAR_INPUT
			dst 	: ^LASCII;
			name 	: ^LASCII;
		END_VAR;

	FUNCTION Free;

	FUNCTION LoadProjectEntries
		VAR_OUTPUT
			retcode 	: BOOL;
		END_VAR;

	FUNCTION ScreenCreate
		VAR_INPUT
			screennumber 	: UDINT;
		END_VAR
		VAR_OUTPUT
			retcode 	: BOOL;
		END_VAR;

	FUNCTION ScreenStart
		VAR_INPUT
			screennumber 	: UDINT;
			startfunct 	: UINT;
			endfunct 	: UINT;
		END_VAR;

	FUNCTION ScreenStop
		VAR_INPUT
			screennumber 	: UDINT;
		END_VAR
		VAR_OUTPUT
			retcode 	: BOOL;
		END_VAR;

	FUNCTION ScreenAddRectangle
		VAR_INPUT
			ptr 	: ^HMI_CTRL_RECTANGLE;
		END_VAR
		VAR_OUTPUT
			retcode 	: BOOL;
		END_VAR;

	FUNCTION ScreenAddLine
		VAR_INPUT
			ptr 	: ^HMI_CTRL_LINE;
		END_VAR
		VAR_OUTPUT
			retcode 	: BOOL;
		END_VAR;

	FUNCTION ScreenAddCtrlImage
		VAR_INPUT
			ptr 	: ^HMI_CTRL_IMAGE;
		END_VAR
		VAR_OUTPUT
			retcode 	: BOOL;
		END_VAR;

	FUNCTION ScreenAddCtrlText
		VAR_INPUT
			ptr 	: ^HMI_CTRL_TEXT;
		END_VAR
		VAR_OUTPUT
			retcode 	: BOOL;
		END_VAR;

	FUNCTION CreateAttrib
		VAR_INPUT
			att32 	: UDINT;
			fontindex 	: UDINT;
		END_VAR
		VAR_OUTPUT
			retcode 	: USINT;
		END_VAR;

	FUNCTION ScreenAddCtrlIO
		VAR_INPUT
			ptr 	: ^HMI_CTRL_IO;
		END_VAR
		VAR_OUTPUT
			retcode 	: BOOL;
		END_VAR;

	FUNCTION AddVariableByName
		VAR_INPUT
			name 	: ^CHAR;
			station 	: UDINT;
		END_VAR
		VAR_OUTPUT
			retcode 	: BOOL;
		END_VAR;

	FUNCTION AddVariable
		VAR_INPUT
			pany 	: ^HMI_ANYTHING;
		END_VAR
		VAR_OUTPUT
			retcode 	: UINT;
		END_VAR;

	FUNCTION AddFont
		VAR_INPUT
			index 	: UDINT;
		END_VAR
		VAR_OUTPUT
			retcode 	: USINT;
		END_VAR;

	FUNCTION AddText
		VAR_INPUT
			pany 	: ^HMI_ANYTHING;
		END_VAR
		VAR_OUTPUT
			retcode 	: UINT;
		END_VAR;

	FUNCTION AddImage
		VAR_INPUT
			pany 	: ^HMI_ANYTHING;
		END_VAR
		VAR_OUTPUT
			retcode 	: UINT;
		END_VAR;

	FUNCTION ScreenAddCtrlRectangle
		VAR_INPUT
			ptr 	: ^HMI_CTRL_RECTANGLE;
		END_VAR
		VAR_OUTPUT
			retcode 	: BOOL;
		END_VAR;

	FUNCTION ScreenAddCtrlLine
		VAR_INPUT
			ptr 	: ^HMI_CTRL_LINE;
		END_VAR
		VAR_OUTPUT
			retcode 	: BOOL;
		END_VAR;

	FUNCTION Create
		VAR_OUTPUT
			retcode 	: BOOL;
		END_VAR;

	FUNCTION SendProject
		VAR_INPUT
			ptr 	: ^void;
		END_VAR
		VAR_OUTPUT
			retcode 	: BOOL;
		END_VAR;

	FUNCTION CreateColor
		VAR_INPUT
			colindex 	: USINT;
		END_VAR
		VAR_OUTPUT
			retcode 	: UINT;
		END_VAR;

	FUNCTION CreateFrame
		VAR_INPUT
			frameindex 	: USINT;
			attrib 	: UDINT;
		END_VAR
		VAR_OUTPUT
			retcode 	: USINT;
		END_VAR;

	FUNCTION AddFunctionBlockIO
		VAR_INPUT
			pany 	: ^HMI_ANYTHING;
		END_VAR
		VAR_OUTPUT
			retcode 	: UINT;
		END_VAR;

	FUNCTION CreateMomStat
		VAR_INPUT
			pio 	: ^HMI_CTRL_IO;
		END_VAR
		VAR_OUTPUT
			retcode 	: UINT;
		END_VAR;

	FUNCTION GLOBAL AddAnything
		VAR_INPUT
			pany 	: ^HMI_ANYTHING;
		END_VAR
		VAR_OUTPUT
			retcode 	: UINT;
		END_VAR;

	FUNCTION AddSheme
		VAR_INPUT
			pany 	: ^HMI_ANYTHING;
		END_VAR
		VAR_OUTPUT
			retcode 	: UINT;
		END_VAR;

	FUNCTION GLOBAL AddFunctionBlock
		VAR_INPUT
			functindex 	: UDINT;
		END_VAR
		VAR_OUTPUT
			retcode 	: UINT;
		END_VAR;

	FUNCTION Run;

	FUNCTION GetFontInfo
		VAR_INPUT
			fontindex 	: UDINT;
		END_VAR
		VAR_OUTPUT
			retcode 	: ^HMI_FONTINFO;
		END_VAR;

	FUNCTION AddImageByIndex
		VAR_INPUT
			index 	: UDINT;
			bootimage 	: BOOL;
		END_VAR
		VAR_OUTPUT
			retcode 	: UINT;
		END_VAR;

	FUNCTION VIRTUAL GLOBAL UpdateValue35
		VAR_INPUT
			varno 	: UINT;
			value 	: DINT;
		END_VAR;

	FUNCTION VIRTUAL GLOBAL UpdateTemperature35
		VAR_INPUT
			value 	: DINT;
		END_VAR;
				//! <Function Comment="method is used to define name of bootimage" Name="GetBootImage"/>
	FUNCTION VIRTUAL GLOBAL GetBootImage
		VAR_OUTPUT
			retcode 	: ^CHAR;
		END_VAR;

	FUNCTION UpLoadProject
		VAR_OUTPUT
			retcode 	: BOOL;
		END_VAR;

	FUNCTION GetVariable
		VAR_INPUT
			pany 	: ^HMI_ANYTHING;
		END_VAR
		VAR_OUTPUT
			retcode 	: ^HMI_VARINFO;
		END_VAR;

	FUNCTION VIRTUAL GLOBAL UpdateString35
		VAR_INPUT
			varno 	: UINT;
			pstr 	: ^void;
			chrsize 	: UDINT;
		END_VAR;

	FUNCTION GLOBAL UpdateAliveSignal35;

	FUNCTION GLOBAL UpdateBacklight35
		VAR_INPUT
			state 	: DINT;
		END_VAR;

	FUNCTION GLOBAL UpdateScreenshot
		VAR_INPUT
			pscrshot 	: ^void;
		END_VAR;

	FUNCTION GLOBAL UpdateActScreen
		VAR_INPUT
			scrno 	: DINT;
		END_VAR;

	FUNCTION GLOBAL UpdateInUse;
				//! <Function Comment="method is used to update firmware in hmi. E:\EasyFirmware.bin&#10; will be used as updatefile." Name="SendNewFirmware"/>
	FUNCTION GLOBAL SendNewFirmware
		VAR_OUTPUT
			retcode 	: BOOL;
		END_VAR;

	FUNCTION GLOBAL OutMessage
		VAR_INPUT
			txt 	: ^CHAR;
		END_VAR;

	FUNCTION GetBacklightDim
		VAR_OUTPUT
			retcode 	: USINT;
		END_VAR;

	FUNCTION OutMessageValue
		VAR_INPUT
			txt 	: ^CHAR;
			value 	: UDINT;
		END_VAR;

	FUNCTION ErrorStateSvr
		VAR_INPUT
			restart 	: BOOL;
		END_VAR;
				//! <Function Comment="method is used to define drive and path of several updatefiles&#13;&#10;note: &quot;E:\&quot; is used as default" Name="GetUpdatePath"/>
	FUNCTION VIRTUAL GLOBAL GetUpdatePath
		VAR_OUTPUT
			retcode 	: ^CHAR;
		END_VAR;
				//! <Function Comment="method is used to define name and location of firmwareupdatefile" Name="GetFirmwareUpdate"/>
	FUNCTION VIRTUAL GLOBAL GetFirmwareUpdate
		VAR_OUTPUT
			retcode 	: ^CHAR;
		END_VAR;
				//! <Function Comment="method is used to define name and location of bootloaderupdatefile" Name="GetBootLoaderUpdate"/>
	FUNCTION VIRTUAL GLOBAL GetBootLoaderUpdate
		VAR_OUTPUT
			retcode 	: ^CHAR;
		END_VAR;
				//! <Function Comment="method will be called once after hmi has (re)started successfully" Name="HmiReady"/>
	FUNCTION VIRTUAL GLOBAL HmiReady;
				//! <Function Comment="methode will be called cyclic when hmi is running" Name="HmiRun"/>
	FUNCTION VIRTUAL GLOBAL HmiRun;

	FUNCTION GetLasalId
		VAR_INPUT
			pany 	: ^HMI_ANYTHING;
		END_VAR
		VAR_OUTPUT
			retcode 	: UDINT;
		END_VAR;

	FUNCTION CreateBarState
		VAR_INPUT
			attrib 	: UDINT;
		END_VAR
		VAR_OUTPUT
			retcode 	: USINT;
		END_VAR;
				//! <Function Comment="method can be used to send multiple data shown in trend at hmi.&#13;&#10;id ....... trendid (0, 1)&#13;&#10;pdata .... pointer to array of trenddata (0 to 255)&#13;&#10;length ... number of valid data in array or 0 to delete actual trenddata in hmi " Name="SendTrend"/>
	FUNCTION GLOBAL SendTrend
		VAR_INPUT
			id 	: UDINT;
			pdata 	: ^USINT;
			length 	: UDINT;
		END_VAR;
				//! <Function Comment="method is used to send pixmap (eg.barcode, qr code) shown at hmi.&#13;&#10;pdata ...... pointer to array of pixmapdata (pitwise pixel)&#13;&#10;width ...... width of pixmap&#13;&#10;height ..... height of pixmap&#13;&#10;padding .... padding (blank) of pixmap&#13;&#10;method will return true on success&#13;&#10;&#13;&#10;to erase pixmap from hmi call methode like SendPixMap(nil, 0, 0, 0);" Name="SendPixMap"/>
	FUNCTION GLOBAL SendPixMap
		VAR_INPUT
			pdata 	: ^void;
			width 	: USINT;
			height 	: USINT;
			padding 	: USINT;
		END_VAR
		VAR_OUTPUT
			retcode 	: BOOL;
		END_VAR;

	FUNCTION GLOBAL UpdateAll
		VAR_INPUT
			act_hmi_crc 	: UDINT;
		END_VAR;

	FUNCTION CheckCrc;

	FUNCTION SleepNext
		VAR_INPUT
			next 	: TStateSvr;
			sleep 	: UDINT;
		END_VAR
		VAR_OUTPUT
			retcode 	: TStateSvr;
		END_VAR;

	FUNCTION SetErrorSvr
		VAR_INPUT
			err 	: TErrorSvr;
		END_VAR;

	FUNCTION CreateVarConst
		VAR_INPUT
			vstate 	: ^USINT;
			pany 	: ^HMI_ANYTHING;
			pdata 	: ^HMI_ANYTHING;
			isog 	: BOOL;
			defval 	: DINT;
		END_VAR
		VAR_OUTPUT
			retcode 	: DINT;
		END_VAR;
				//! <Function Comment="methode is used to ask for actual access by using accesslevel" Name="HmiAccess"/>
	FUNCTION VIRTUAL GLOBAL HmiAccess
		VAR_INPUT
			level 	: UDINT;			//! <Variable Comment="accesslevel" Name="HmiAccess.level"/>
		END_VAR
		VAR_OUTPUT
			retcode 	: BOOL;			//! <Variable Comment="return true if access is given&#13;&#10;on the other hand return false (writeprotected)" Name="HmiAccess.retcode"/>
		END_VAR;

	FUNCTION GLOBAL SoftResetAll;

	FUNCTION GLOBAL SoftReset;

	FUNCTION ScreenAddCtrlCircle
		VAR_INPUT
			ptr 	: ^HMI_CTRL_CIRCLE;
		END_VAR
		VAR_OUTPUT
			retcode 	: BOOL;
		END_VAR;

	FUNCTION GetEnumSchemeIndex
		VAR_INPUT
			pany 	: ^HMI_ANYTHING;
		END_VAR
		VAR_OUTPUT
			retcode 	: UDINT;
		END_VAR;
				//! <Function Comment="method is used to perform defined &quot;UserCall&quot;. overwrite method to implement userspecific code by using parameter" Name="UserCall"/>
	FUNCTION VIRTUAL GLOBAL UserCall
		VAR_INPUT
			fktno 	: UDINT;
			para 	: DINT;
		END_VAR;

	FUNCTION CheckProjectCrc
		VAR_INPUT
			ptr 	: ^void;
			hmiver 	: UDINT;
			chkold 	: BOOL;
		END_VAR
		VAR_OUTPUT
			retcode 	: BOOL;
		END_VAR;
				//! <Function Comment="method is used to add some text, image, variables, etc. to project sent to hmi before lse-project is added" Name="HmiProjectBegin"/>
	FUNCTION VIRTUAL GLOBAL HmiProjectBegin;
				//! <Function Comment="method is used to add some text, image, etc. to project sent to hmi" Name="HmiProjectCreate"/>
	FUNCTION VIRTUAL GLOBAL HmiProjectCreate;
				//! <Function Comment="method can be used to add userdefined text to project sent to hmi.&#13;&#10;the id of added text will be returned.&#13;&#10;note: method has to be called in overwritten virtual method HmiProjectCreate()" Name="CreateAddText"/>
	FUNCTION CreateAddText
		VAR_INPUT
			txt 	: ^void;
			chrsize 	: UDINT;
		END_VAR
		VAR_OUTPUT
			retcode 	: UDINT;
		END_VAR;
				//! <Function Comment="method can be used to add new image to project sent to hmi.&#13;&#10;the id of added image will be returned.&#13;&#10;note: method has to be called in oerwritten virtual method HmiProjectCreate()" Name="CreateAddImage"/>
	FUNCTION CreateAddImage
		VAR_INPUT
			txt 	: ^CHAR;
		END_VAR
		VAR_OUTPUT
			retcode 	: UDINT;
		END_VAR;
				//! <Function Comment="method is used to customise listcontrol at hmi&#13;&#10;listid ............ id of list to customise (0)&#13;&#10;lineno_max ........ max. number of lstitems in list&#13;&#10;line_height ....... height of listitem in pixel&#13;&#10;items_per_line .... number of listitems shown in each line&#13;&#10;datim2line ........ view date and time next(false) or on top(true) to each other&#13;&#10;bottom_up ...... view last line always on top (Firmwareversion &gt;= 1.48 needed)&#13;&#10;&#13;&#10;" Name="ListSetup"/>
	FUNCTION GLOBAL ListSetup
		VAR_INPUT
			listid 	: UDINT;
			lineno_max 	: UDINT;
			line_height 	: UDINT;
			items_per_line 	: UDINT;
			datim2line 	: BOOL;
			bottom_up 	: BOOL := false;
		END_VAR
		VAR_OUTPUT
			retcode 	: BOOL;
		END_VAR;
				//! <Function Comment="method is used to send some commands to listcontrol at hmi&#13;&#10;listid ............ id of list to customise (0)&#13;&#10;cmd ............... 0...delete all items of listcontrol&#13;&#10;                    1...deselect actual selected item&#13;&#10;                    2...delete single item in list &#13;&#10;item_index ........ is used to address item&#13;&#10;&#13;&#10;" Name="ListCmd"/>
	FUNCTION GLOBAL ListCmd
		VAR_INPUT
			listid 	: UDINT;
			cmd 	: UDINT;
			item_index 	: UDINT;
		END_VAR
		VAR_OUTPUT
			retcode 	: BOOL;
		END_VAR;
				//! <Function Comment="method is used to add item to listcontrol at hmi. listcontrol will act as ringbuffer with 200 entries.&#13;&#10;listid ............ id of list to customise (0)&#13;&#10;item_type ......... 2...text&#13;&#10;                    3...image&#13;&#10;item_val ........... index of text or image&#13;&#10;item_date ......... date of itementry or 0&#13;&#10;item_time ......... time of itementry or 0&#13;&#10;if &quot;item_date&quot; and &quot;item_time&quot; are set to 0, no information about date and time will be shown at item in hmi.&#13;&#10;" Name="ListAddEntry"/>
	FUNCTION GLOBAL ListAddEntry
		VAR_INPUT
			listid 	: UDINT;
			item_type 	: UDINT;
			item_val 	: UDINT;
			item_date 	: UDINT;
			item_time 	: UDINT;
		END_VAR
		VAR_OUTPUT
			retcode 	: BOOL;
		END_VAR;
				//! <Function Comment="method is used to add some deeds to actual processed screen sent to hmi&#13;&#10;screenno .... number of screen in process" Name="HmiScreenCreate"/>
	FUNCTION VIRTUAL GLOBAL HmiScreenCreate
		VAR_INPUT
			screenno 	: UDINT;
		END_VAR;
				//! <Function Comment="method is used to indicate if english format of date (&quot;month/day/year&quot;) and time (&quot;01:30.10pm&quot;) is in use (retcode:=true).&#13;&#10;otherwise (retcode:=false) date will be represented as &quot;day.month.year&quot; and time as &quot;13:30:10&quot;" Name="EnglishFormatDateTime"/>
	FUNCTION VIRTUAL GLOBAL EnglishFormatDateTime
		VAR_INPUT
			languageid 	: UDINT;
		END_VAR
		VAR_OUTPUT
			retcode 	: BOOL;
		END_VAR;
				//! <Function Comment="method is used to define number of &quot;userextended variables&quot; done in firmware of hmi" Name="HmiVariableExtention"/>
	FUNCTION VIRTUAL GLOBAL HmiVariableExtention
		VAR_INPUT
			varname 	: ^CHAR;
		END_VAR
		VAR_OUTPUT
			retcode 	: UDINT;
		END_VAR;

	FUNCTION VIRTUAL IsProjectUpLoadNecessary
		VAR_INPUT
			preselect 	: BOOL;
		END_VAR
		VAR_OUTPUT
			retcode 	: BOOL;
		END_VAR;
				//! <Function Comment="method is used to create crc including all dynamic parts (without ststic data) from hmi-project.&#13;&#10;call method (get crc) in derived method IsProjectUpLoadNecessary() " Name="GetMapCrc"/>
	FUNCTION GetMapCrc
		VAR_OUTPUT
			retcode 	: UDINT;
		END_VAR;

	FUNCTION VIRTUAL GLOBAL UpdatePixMap
		VAR_INPUT
			value 	: DINT;
		END_VAR
		VAR_OUTPUT
			retcode 	: DINT;
		END_VAR;

	FUNCTION VIRTUAL GLOBAL UpdateTrendVal
		VAR_INPUT
			id 	: UDINT;
			value 	: DINT;
		END_VAR
		VAR_OUTPUT
			retcode 	: DINT;
		END_VAR;
				//! <Function Comment="method is used to recalculate binary-values to physical-values in both directions&#13;&#10;value ....... actual value&#13;&#10;formula ..... information about used physcal formula&#13;&#10;dezpoint .... number of digits on right side of decimalpoint&#13;&#10;direction ... true = sps--&gt;hmi (binary to physic), false = hmi--&gt;sps (physic to binary)" Name="Recalculate"/>
	FUNCTION VIRTUAL GLOBAL Recalculate
		VAR_INPUT
			value 	: DINT;
			formula 	: UDINT;
			dezpoint 	: DINT;
			direction 	: BOOL;
		END_VAR
		VAR_OUTPUT
			retcode 	: DINT;
		END_VAR;

	FUNCTION VIRTUAL IsProjectUpLoadNecessaryEx
		VAR_INPUT
			preselect 	: BOOL;
			crc_hmi 	: UDINT;			//! <Variable Comment="actual crc got from HMI. 0 ... no connection to HMI, 0xFFFFFFFF ... no project in HMI, any other value is valid crc" Name="IsProjectUpLoadNecessaryEx.crc_hmi"/>
			crc_prj 	: UDINT;			//! <Variable Comment="actual crc computed in plc" Name="IsProjectUpLoadNecessaryEx.crc_prj"/>
		END_VAR
		VAR_OUTPUT
			retcode 	: BOOL;			//! <Variable Comment="return &apos;true&apos; to upload project to HMI, on the other hand return &apos;false&apos;" Name="IsProjectUpLoadNecessaryEx.retcode"/>
		END_VAR;

	FUNCTION VIRTUAL Recalculate_Stroke2mm
		VAR_INPUT
			value 	: DINT;
			dezpoint 	: DINT;
			direction 	: BOOL;
		END_VAR
		VAR_OUTPUT
			retcode 	: DINT;
		END_VAR;

	FUNCTION VIRTUAL Recalculate_Stroke2inch
		VAR_INPUT
			value 	: DINT;
			dezpoint 	: DINT;
			direction 	: BOOL;
		END_VAR
		VAR_OUTPUT
			retcode 	: DINT;
		END_VAR;

	FUNCTION Recalculate_MulDiv
		VAR_INPUT
			einheit 	: UDINT;
			posdezpt 	: DINT;
		END_VAR
		VAR_OUTPUT
			retcode 	: DINT;
		END_VAR;

	FUNCTION VIRTUAL Recalculate_Temp2Celsius
		VAR_INPUT
			value 	: DINT;
			dezpoint 	: DINT;
			direction 	: BOOL;
		END_VAR
		VAR_OUTPUT
			retcode 	: DINT;
		END_VAR;

	FUNCTION VIRTUAL Recalculate_Temp2Fahrenheit
		VAR_INPUT
			value 	: DINT;
			dezpoint 	: DINT;
			direction 	: BOOL;
		END_VAR
		VAR_OUTPUT
			retcode 	: DINT;
		END_VAR;

	FUNCTION VIRTUAL Recalculate_Weight2Kilogram
		VAR_INPUT
			value 	: DINT;
			dezpoint 	: DINT;
			direction 	: BOOL;
		END_VAR
		VAR_OUTPUT
			retcode 	: DINT;
		END_VAR;

	FUNCTION VIRTUAL Recalculate_Weight2Pound
		VAR_INPUT
			value 	: DINT;
			dezpoint 	: DINT;
			direction 	: BOOL;
		END_VAR
		VAR_OUTPUT
			retcode 	: DINT;
		END_VAR;

	FUNCTION VIRTUAL Recalculate_Pressure2Bar
		VAR_INPUT
			value 	: DINT;
			dezpoint 	: DINT;
			direction 	: BOOL;
		END_VAR
		VAR_OUTPUT
			retcode 	: DINT;
		END_VAR;

	FUNCTION VIRTUAL Recalculate_Pressure2Psi
		VAR_INPUT
			value 	: DINT;
			dezpoint 	: DINT;
			direction 	: BOOL;
		END_VAR
		VAR_OUTPUT
			retcode 	: DINT;
		END_VAR;

	FUNCTION VIRTUAL Recalculate_Time2Second
		VAR_INPUT
			value 	: DINT;
			dezpoint 	: DINT;
			direction 	: BOOL;
		END_VAR
		VAR_OUTPUT
			retcode 	: DINT;
		END_VAR;

	FUNCTION VIRTUAL Recalculate_Time2Minute
		VAR_INPUT
			value 	: DINT;
			dezpoint 	: DINT;
			direction 	: BOOL;
		END_VAR
		VAR_OUTPUT
			retcode 	: DINT;
		END_VAR;

	FUNCTION VIRTUAL Recalculate_Time2Hour
		VAR_INPUT
			value 	: DINT;
			dezpoint 	: DINT;
			direction 	: BOOL;
		END_VAR
		VAR_OUTPUT
			retcode 	: DINT;
		END_VAR;

	FUNCTION VIRTUAL Recalculate_Force2KN
		VAR_INPUT
			value 	: DINT;
			dezpoint 	: DINT;
			direction 	: BOOL;
		END_VAR
		VAR_OUTPUT
			retcode 	: DINT;
		END_VAR;

	FUNCTION Recalculate_Calc
		VAR_INPUT
			rval 	: REAL;
			rmul 	: REAL;
			rdiv 	: REAL;
			direction 	: BOOL;
		END_VAR
		VAR_OUTPUT
			retcode 	: DINT;
		END_VAR;
				//! <Function Comment="method is used to add some customized text to list&#13;&#10;listid ............ id of list to customise (0/1)&#13;&#10;item_date ......... date of itementry or 0&#13;&#10;item_time ......... time of itementry or 0&#13;&#10;ptxt ..... Pointer to userspezific text&#13;&#10;chrsize ..... Format of userspezific text (1 ... ASCII, 2 ... Unicode)&#13;&#10;item_id ..... individual id of text&#13;&#10;&#13;&#10;" Name="ListAddText"/>
	FUNCTION GLOBAL ListAddText
		VAR_INPUT
			listid 	: UDINT;
			item_date 	: UDINT;
			item_time 	: UDINT;
			ptxt 	: ^void;
			chrsize 	: UDINT;
			item_id 	: UDINT;
		END_VAR
		VAR_OUTPUT
			retcode 	: BOOL;
		END_VAR;

	FUNCTION GLOBAL SoftResetIn
		VAR_INPUT
			milliseconds 	: UDINT;
		END_VAR;
				//! <Function Comment="method will be called each time when ir-code is detected on hmi.&#13;&#10;code ... detected code&#13;&#10;note: functionality is just given when hmi supports ir-detection" Name="UpdateIrCode"/>
	FUNCTION VIRTUAL UpdateIrCode
		VAR_INPUT
			code 	: UDINT;
		END_VAR;

	FUNCTION SendUpdateToHmi
		VAR_INPUT
			dpne 	: ^CHAR;
		END_VAR
		VAR_OUTPUT
			retcode 	: BOOL;
		END_VAR;

	FUNCTION GLOBAL SendNewBootLoader
		VAR_OUTPUT
			retcode 	: BOOL;
		END_VAR;

	FUNCTION VIRTUAL GLOBAL CheckUpdate
		VAR_INPUT
			dpne 	: ^CHAR;
			nextstep 	: TStateSvr;
			defaultstep 	: TStateSvr;
			sleep 	: UDINT;
		END_VAR
		VAR_OUTPUT
			retcode 	: TStateSvr;
		END_VAR;
				//! <Function Comment="Get NoticeText from lse-project. &#13;&#10;Method will return pointer to ascii-0-string or NIL if NoticeText is empty." Name="GetLseProjectNotice"/>
	FUNCTION GLOBAL GetLseProjectNotice
		VAR_OUTPUT
			retcode 	: ^CHAR;
		END_VAR;
				//! <Function Comment="User is able to set RevisionNumber of HMI-Software by using this method." Name="UserProjectRevision"/>
	FUNCTION VIRTUAL GLOBAL UserProjectRevision
		VAR_OUTPUT
			retcode 	: UINT;
		END_VAR;

	FUNCTION AddStateBitByName
		VAR_INPUT
			name 	: ^CHAR;
			invert 	: BOOL;
			access 	: UINT;
		END_VAR
		VAR_OUTPUT
			retcode 	: BOOL;
		END_VAR;

	FUNCTION SaveFile
		VAR_INPUT
			dp 	: ^CHAR;
			fileid 	: UDINT;
			size 	: UDINT;
			ptr 	: ^void;
		END_VAR
		VAR_OUTPUT
			retcode 	: BOOL;
		END_VAR;

	FUNCTION SaveProject
		VAR_INPUT
			dp 	: ^CHAR;
			prj 	: ^void;
		END_VAR;
				//! <Function Comment="use methode to enable variable Limits at HMI.&#13;&#10;retcode = false .... limits at Variables are static&#13;&#10;retcode = true .... variable limits at Variables will work&#13;&#10;" Name="VariableLimitsInUse"/>
	FUNCTION VIRTUAL GLOBAL VariableLimitsInUse
		VAR_OUTPUT
			retcode 	: DINT;
		END_VAR;

	FUNCTION GetObjectName
		VAR_INPUT
			pthis 	: ^void;
		END_VAR
		VAR_OUTPUT
			retcode 	: ^CHAR;
		END_VAR;

	FUNCTION VIRTUAL GLOBAL UpdateHumidity35
		VAR_INPUT
			value 	: DINT;
		END_VAR;
				//! <Function Comment="Method can be used (overwrite) to change name of individual Object or use OverloadLight mechanism at default" Name="HmiOverloadLight"/>
	FUNCTION VIRTUAL GLOBAL HmiOverloadLight;

	FUNCTION ListAddEntryIntern
		VAR_INPUT
			listid 	: UDINT;
			item_type 	: UDINT;
			item_val 	: UDINT;
			item_date 	: UDINT;
			item_time 	: UDINT;
			ptxt 	: ^void;
			chrsize 	: UDINT;
			item_id 	: UDINT;
		END_VAR
		VAR_OUTPUT
			retcode 	: BOOL;
		END_VAR;
				//! <Function Comment="Get copy of Lse-project-name. " Name="GetLseProjectName"/>
	FUNCTION GLOBAL GetLseProjectName
		VAR_INPUT
			pdst 	: ^void;			//! <Variable Comment="Pointer to destination where projectname should be filed" Name="GetLseProjectName.pdst"/>
			dchrsize 	: UDINT;			//! <Variable Comment="Bytesize of single character to be filed (1..Ascii, 2..Unicode)" Name="GetLseProjectName.dchrsize"/>
			bytesize_dst 	: UDINT;			//! <Variable Comment="Bytesize of destination. Note: Destination has to be big enought to cover name, otherwise name will be truncated." Name="GetLseProjectName.bytesize_dst"/>
		END_VAR;
				//! <Function Comment="Method can be used to configurate T9-Keypad at HMI.&#13;&#10;Note: Firmware 1.46 or greater is needed at HMI, otherwise configuration will be ignored." Name="T9KeyboardConfig"/>
	FUNCTION VIRTUAL GLOBAL T9KeyboardConfig;

	FUNCTION VIRTUAL GLOBAL ClassSvr::NewInst
		VAR_INPUT
			pPara 	: ^CmdStruct;
			pResult 	: ^results;
		END_VAR
		VAR_OUTPUT
			ret_code 	: iprStates;
		END_VAR;

	FUNCTION VIRTUAL GLOBAL StateSvr::Write
		VAR_INPUT
			input (EAX) 	: LseEasy::TStateSvr;
		END_VAR
		VAR_OUTPUT
			result (EAX) 	: LseEasy::TStateSvr;
		END_VAR;

	FUNCTION VIRTUAL GLOBAL ActLanguage::Write
		VAR_INPUT
			input (EAX) 	: UDINT;
		END_VAR
		VAR_OUTPUT
			result (EAX) 	: UDINT;
		END_VAR;

	FUNCTION VIRTUAL GLOBAL ActScreen::Write
		VAR_INPUT
			input (EAX) 	: DINT;
		END_VAR
		VAR_OUTPUT
			result (EAX) 	: DINT;
		END_VAR;

	FUNCTION VIRTUAL GLOBAL BacklightOnOff::Write
		VAR_INPUT
			input (EAX) 	: DINT;
		END_VAR
		VAR_OUTPUT
			result (EAX) 	: DINT;
		END_VAR;

	FUNCTION VIRTUAL GLOBAL BacklightDim::Write
		VAR_INPUT
			input (EAX) 	: DINT;
		END_VAR
		VAR_OUTPUT
			result (EAX) 	: DINT;
		END_VAR;
  //Tables:
	FUNCTION @STD
		VAR_OUTPUT
			ret_code	: CONFSTATES;
		END_VAR;
	FUNCTION GLOBAL TAB @CT_;
END_CLASS;

#pragma using HmiChkBitList
#pragma using HmiColorMap
#pragma using HmiFile
#pragma using HmiFont35
#pragma using HmiFontList
#pragma using HmiFunctionList
#pragma using HmiFunctionList35
#pragma using HmiImage35
#pragma using HmiImageList
#pragma using HmiMapFile
#pragma using HmiProject35
#pragma using HmiProjectList
#pragma using HmiScreen
#pragma using HmiSetUpList
#pragma using HmiSetupList35
#pragma using HmiShemeList
#pragma using HmiShemeList35
#pragma using HmiStateBit35
#pragma using HmiStrLib
#pragma using HmiT9Config35
#pragma using HmiTextList
#pragma using HmiTextList35
#pragma using HmiUtils
#pragma using HmiVarList
#pragma using HmiVarList35
#pragma usingLtd HmiComPort

#includeC "..\LseEasy\Create.h"

#define DEFAULT_VALUE_HUMIDITY    -32768
#define DEFAULT_VALUE_TEMPERATURE -32768
#define FUEHLERBRUCH              16#80000010

var_private
  InstanceCnt : UDINT;
  InstancePtr : Array[0..31] of ^LseEasy;
end_var

FUNCTION LseEasy::LseEasy
	VAR_OUTPUT
		ret_code 	: ConfStates;
	END_VAR

  InstanceCnt   := 0;
	ret_code      := C_OK;
  StateSvr      := TStart;
  ProjectBox    := nil;
  HmiPrjCrc     := 1; // has to be set to 1 !!
  Hmi35PrjCrc   := 0; // has to be set to 0 !!
  TryToRestart  := false;
  CallScreen    := -1;
  ActScreen     := -1;
  TrendVal0     := -1;
  TrendVal1     := -1;
  ListVal0      := -1;
  ListVal1      := -1;
  PixMap        := -1;
  NeedUpdateAll := 0;
  AutoFwUpdateDisabled := false;
  ActTemperature := DEFAULT_VALUE_TEMPERATURE;
  ActHumidity    := DEFAULT_VALUE_HUMIDITY;

END_FUNCTION

FUNCTION VIRTUAL GLOBAL LseEasy::Init
  VAR
  	ph : ^dint;
  END_VAR

  ph := (#ListVal0) - 4;
  ListVal0Lid := ph$udint;
  ph := (#ListVal1) - 4;
  ListVal1Lid := ph$udint;
  ph := (#TrendVal0) - 4;
  TrendVal0Lid := ph$udint;
  ph := (#TrendVal1) - 4;
  TrendVal1Lid := ph$udint;
  ph := (#BacklightDim) - 4;
  BacklightDimLid := ph$udint;
  ph := (#HmiSwVersion) - 4;
  HmiSwVersionLid := ph$udint;
  ph := (#HmiHwVersion) - 4;
  HmiHwVersionLid := ph$udint;
  ph := (#PixMap) - 4;
  PixMapLid       := ph$udint;

  if(_FirstScan) then
    if(InstanceCnt < (sizeof(InstancePtr) / sizeof(InstancePtr[0]))) then
      InstancePtr[InstanceCnt] := this;
      InstanceCnt += 1;
    end_if;
    ComPort.Start(this);
    HmiVarList.SetSuper(this);
  end_if;

END_FUNCTION

FUNCTION LseEasy::Free

  HmiPrjCrc     := 1; // has to be set to 1 !!
  Hmi35PrjCrc   := 0; // has to be set to 0 !!
  ProjectBox    := nil;
  RefreshTix    := 0;
  TrendVal0     := -1;
  TrendVal1     := -1;
  ListVal0      := -1;
  ListVal1      := -1;
  PixMap        := -1;
  LastUsage     := 0;
  NeedUpdateAll := 1;
  HmiOnline     := 0; // hmi is offline
  CantGetCrc    := 0;
  ErrorSvr      := ErrNone;
  HmiSwVersion  := 0;
  HmiHwVersion  := 0;
  ActTemperature := DEFAULT_VALUE_TEMPERATURE;
  ActHumidity    := DEFAULT_VALUE_HUMIDITY;

END_FUNCTION

FUNCTION LseEasy::SetErrorSvr
	VAR_INPUT
		err 	: TErrorSvr;
	END_VAR

  if(ErrorSvr = ErrNone) then
    ErrorSvr := err;
  end_if;

END_FUNCTION

FUNCTION LseEasy::GetObjectName
	VAR_INPUT
    pthis : ^void;
  END_VAR
  VAR_OUTPUT
    retcode : ^char;
  END_VAR
  VAR
  	pobj : ^OBJ;
  END_VAR

  pobj$^void := pthis;
  pobj -= sizeof(OBJ);
  retcode$^CLexem := #pobj^.pObjDsc^.SymName;
  retcode += 4;

END_FUNCTION

FUNCTION VIRTUAL GLOBAL LseEasy::GetPrjPath
	VAR_OUTPUT
		retcode 	: ^LASCII;
	END_VAR

  ProjectPath := ProjectPath.Read();

  if(ProjectPath > 0) then // SA42417
    StringLib.StrCpy(#LseProjectPath[0], 1, "C:\Easy", 1);
    StringLib.DintToStr(#LseProjectPath[7], ProjectPath, 16#800, 1);
    StringLib.StrCat(#LseProjectPath[0], 1, "\", 1);
  elsif(ProjectPath = -1) then // SA42417
    StringLib.StrCpy(#LseProjectPath[0], 1, "C:\", 1);
    StringLib.StrCat(#LseProjectPath[0], 1, GetObjectName(this), 1);
    StringLib.StrCat(#LseProjectPath[0], 1, "\", 1);
  else
    StringLib.StrCpy(#LseProjectPath[0], 1, "C:\MPC\", 1);
  end_if;

  retcode := #LseProjectPath[0];

END_FUNCTION

FUNCTION VIRTUAL GLOBAL LseEasy::GetBootImage
	VAR_OUTPUT
		retcode 	: ^CHAR;
	END_VAR

  retcode := "bootimage"; // name of bootimage

END_FUNCTION

FUNCTION VIRTUAL GLOBAL LseEasy::GetUpdatePath
	VAR_OUTPUT
		retcode 	: ^CHAR;
	END_VAR

  retcode := "E:\";

END_FUNCTION

FUNCTION VIRTUAL GLOBAL LseEasy::GetFirmwareUpdate
	VAR_OUTPUT
		retcode 	: ^CHAR;
	END_VAR

  StringLib.StrCpy(#UpdateFileDPNE[0], 1, GetUpdatePath(), 1);
  StringLib.StrCat(#UpdateFileDPNE[0], 1, "EasyFirmware.bin", 1);
  retcode := #UpdateFileDPNE[0]; // drive:\path\name.extention of firmwareupdatefile

END_FUNCTION

FUNCTION VIRTUAL GLOBAL LseEasy::GetBootLoaderUpdate
	VAR_OUTPUT
		retcode 	: ^CHAR;
	END_VAR

  StringLib.StrCpy(#UpdateFileDPNE[0], 1, GetUpdatePath(), 1);
  StringLib.StrCat(#UpdateFileDPNE[0], 1, "BootKiller.bin", 1);
  retcode := #UpdateFileDPNE[0]; // drive:\path\name.extention of bootloaderupdatefile

END_FUNCTION

FUNCTION VIRTUAL GLOBAL LseEasy::HmiReady

END_FUNCTION

FUNCTION VIRTUAL GLOBAL LseEasy::HmiRun
//  VAR
//  	vno : udint;
//    txt : array[0..100] of char;
//  END_VAR
//
//  vno := HmiVarList.GetVarNoByName("Dummy.Server2", 0);
//  HmiVarList.GetServerName(#txt[0], vno);

END_FUNCTION

FUNCTION VIRTUAL GLOBAL LseEasy::HmiOverloadLight
  VAR
  	ovl : dint;
  END_VAR

  ovl := OverloadLight.Read();
  HmiVarList.OverloadLight(ovl);

//  case ovl of
//    1 : HmiVarList.RenameRootObject("Dummy", "LivingRoom");
//    2 : HmiVarList.RenameRootObject("Dummy", "BathRoom");
//    3 : HmiVarList.RenameRootObject("Dummy", "Office");
//  end_case;

END_FUNCTION

FUNCTION VIRTUAL GLOBAL LseEasy::VariableLimitsInUse
	VAR_OUTPUT
		retcode 	: DINT;
	END_VAR

  retcode := false; // don't use variable limits at Server

END_FUNCTION

FUNCTION LseEasy::ErrorStateSvr
  VAR_INPUT
    restart : bool;
  END_VAR

  StateSvr          := TError;
  AliveTix35CntrOld := AliveTix35Cntr;
  TryToRestart      := restart;

END_FUNCTION

FUNCTION LseEasy::SleepNext
	VAR_INPUT
		next 	: TStateSvr;
		sleep 	: UDINT;
	END_VAR
	VAR_OUTPUT
		retcode 	: TStateSvr;
	END_VAR

  StateSvr      := TSleep;
  StateNext     := next;
  SleepStart    := ops.tAbsolute;
  SleepDuration := sleep;
  retcode       := StateSvr;

END_FUNCTION

FUNCTION LseEasy::MakePrjFileName
	VAR_INPUT
		dst 	: ^LASCII;
		name 	: ^LASCII;
	END_VAR

  StringLib.StrCpy(dst, sizeof(char), GetPrjPath(), sizeof(char));
  StringLib.StrCat(dst, sizeof(char), name, sizeof(char));

END_FUNCTION

FUNCTION LseEasy::UpLoadProject
	VAR_OUTPUT
		retcode 	: BOOL;
	END_VAR

  retcode := false;

  if(ProjectBox <> NIL) then
    if(SendProject(ProjectBox) = true) then
      retcode := true;
    else
      ErrorStateSvr(true);
    end_if;
  end_if;

END_FUNCTION

FUNCTION LseEasy::CreateAddText
	VAR_INPUT
    txt : ^void;
    chrsize : udint;
	END_VAR
	VAR_OUTPUT
		retcode 	: udint;
	END_VAR
  VAR
  	tmp : array[0..255] of uint;
    pa : ^usint;
    pu : ^uint;
  END_VAR

  retcode := 16#FFFFFFFF;
  if((CreateAdd = true) & (txt <> NIL)) then
    if(chrsize = 1) then
      pa := txt$^usint;
      pu := #tmp[0];
      while(pa^) do
        pu^ := pa^;
        pu += 2;
        pa += 1;
      end_while;

      pu^ := 0;
      txt$^uint := #tmp[0];
    end_if;
    retcode := HmiTextList35.AddEntry(txt$^uint);
  end_if;

END_FUNCTION

FUNCTION LseEasy::CreateAddImage
	VAR_INPUT
    txt : ^char;
	END_VAR
	VAR_OUTPUT
		retcode 	: udint;
	END_VAR

  retcode := 16#FFFFFFFF;
  if((CreateAdd = true) & (txt <> NIL)) then
    retcode := AddImageByIndex(HmiImageList.GetIndexByName(txt), false);
  end_if;

END_FUNCTION

FUNCTION GLOBAL LseEasy::ListSetup
	VAR_INPUT
		listid 	: UDINT;
		lineno_max 	: UDINT;
		line_height 	: UDINT;
		items_per_line 	: UDINT;
		datim2line 	: BOOL;
		bottom_up 	: BOOL;(* := false *)
	END_VAR
	VAR_OUTPUT
		retcode 	: BOOL;
	END_VAR
  var
    tmp : array[0..6] of usint;
  end_var

  if(lineno_max > 255) then
    lineno_max := 255;
   end_if;

  retcode := false;
  tmp[0] := ComCMD_UPDATELIST0_CMD;
  if(listid = 0) then // sonderfall, aus kompatibilitätsgründen zu älterer firmware beibehalten
    tmp[1] := 16#FF; // setup
  else
    tmp[1] := (listid$usint shl 4) or 16#0F; // listid + setup
  end_if;

  tmp[2] := items_per_line$usint;
  tmp[3] := line_height$usint;
  tmp[4] := 0;
  if(datim2line = true) then
    tmp[4] := tmp[4] or 1;
  end_if;

  if(HmiSwVersion >= 148) then
    if(bottom_up = true) then
      tmp[4] := tmp[4] or 2;
    end_if;
  end_if;

  tmp[5] := lineno_max$usint;
  tmp[6] := 0; // nc
  retcode := ComPort.SendData(#tmp[0], 7);

END_FUNCTION

FUNCTION GLOBAL LseEasy::ListCmd
	VAR_INPUT
		listid 	: UDINT;
		cmd 	: UDINT;
		item_index 	: UDINT;
	END_VAR
	VAR_OUTPUT
		retcode 	: BOOL;
	END_VAR
  var
    tmp : array[0..6] of usint;
  end_var

  tmp[0]       := ComCMD_UPDATELIST0_CMD;
  tmp[1]       := (listid$usint shl 4) or cmd$usint;
  tmp[2]$udint := item_index;
  tmp[6]       := 0; // nc
  retcode      := ComPort.SendData(#tmp[0], 7);

END_FUNCTION

FUNCTION LseEasy::ListAddEntryIntern
	VAR_INPUT
		listid 	: UDINT;
		item_type 	: UDINT;
		item_val 	: UDINT;
		item_date 	: UDINT;
		item_time 	: UDINT;
		ptxt 	: ^void;
		chrsize 	: UDINT;
		item_id 	: UDINT;
	END_VAR
	VAR_OUTPUT
		retcode 	: BOOL;
	END_VAR
  var
    tmp : array[0..99] of usint;
    datim, tmp32 : udint;
    len, nox : udint;
  end_var

  // -----------TTTTTTOOOOSSSSSMMMMMM
  //                           ||||||
  //                           ++++++ ----- minuten (6 bit)
  //                      +++++ ----------- stunden (5 bit)
  //                  ++++ ---------------- monat (4 bit)
  //            ++++++ -------------------- tag (6 bit)
  // +++++++++++ -------------------------- 0

  // itemtype  1...variable, 2...text, 3...image
  retcode := false;
  if(listid < 2) then

    datim := 0;
    if((item_date <> 0) | (item_time <> 0)) then
      // YYYYYYYYYYYYYYYYMMMMDDDDDDDDWWWW
      // HHHHHHHHNNNNNNNNSSSSSSSSxxxxxxxx
      datim := (item_time shr 16) and 16#3F;
      tmp32 := (item_time shr 24) and 16#1F;
      datim := datim or (tmp32 shl 6);
      tmp32 := (item_date shr 12) and 16#0F;
      datim := datim or (tmp32 shl (6+5));
      tmp32 := (item_date shr 4) and 16#3F;
      datim := datim or (tmp32 shl (6+5+4));
    end_if;

    tmp[0]       := ComCMD_UPDATELIST0_ADD;
    if(listid = 1) then
      tmp[0]     := ComCMD_UPDATELIST1_ADD;
    end_if;
    tmp[1]$uint  := item_val$uint;
    tmp[3]       := item_type$usint;
    tmp[4]$udint := datim;

    len := 7;

    if((item_id <> 16#FFFFFFFF) | (ptxt <> nil)) then
      tmp[7]$udint := item_id;
      len := 11;
    end_if;

    if(ptxt <> nil) then
      if(chrsize > 1) then
        nox := StringLib.StrLen(ptxt, 2);
        if(nox >= 40) then
          nox := 39;
        end_if;
        nox := nox * 2;
        _memcpy(#tmp[len], ptxt, nox);
        len += nox;
        tmp[len]$uint := 0;
        len += 2;
      else
        nox := StringLib.StrLen(ptxt, 1);
        if(nox >= 80) then
          nox := 79;
        end_if;
        _memcpy(#tmp[len], ptxt, nox);
        len += nox;
        tmp[len] := 0;
        len += 1;
      end_if;
    end_if;

    retcode := ComPort.SendData(#tmp[0], len);
  end_if;

END_FUNCTION

FUNCTION GLOBAL LseEasy::ListAddEntry
	VAR_INPUT
		listid 	: UDINT;
		item_type 	: UDINT;
		item_val 	: UDINT;
		item_date 	: UDINT;
		item_time 	: UDINT;
	END_VAR
	VAR_OUTPUT
		retcode 	: BOOL;
	END_VAR

  retcode := ListAddEntryIntern(listid, item_type, item_val, item_date, item_time, nil, 0, 16#FFFFFFFF);

END_FUNCTION

FUNCTION GLOBAL LseEasy::ListAddText
	VAR_INPUT
		listid 	: UDINT;
		item_date 	: UDINT;
		item_time 	: UDINT;
		ptxt 	: ^void;
		chrsize 	: UDINT;
		item_id 	: UDINT;
	END_VAR
	VAR_OUTPUT
		retcode 	: BOOL;
	END_VAR
  VAR
  	item_type : udint;
  END_VAR

  item_type := 4;
  if(chrsize > 1) then
    item_type := 5;
    chrsize := 2;
  end_if;

  retcode := ListAddEntryIntern(listid, item_type, 0, item_date, item_time, ptxt, chrsize, item_id);

END_FUNCTION

FUNCTION VIRTUAL GLOBAL LseEasy::HmiProjectBegin

// AddVariableByName("Objekt.Server", 0); // fix variablennumber in hmi
// AddStateBitByName("CheckBit2", false, 0); // fix statebitnumber in hmi

//  HmiImageList.XChange("spiderman", "E:\Image0.bmp");

END_FUNCTION

FUNCTION VIRTUAL GLOBAL LseEasy::HmiProjectCreate

END_FUNCTION

FUNCTION VIRTUAL GLOBAL LseEasy::UserProjectRevision
	VAR_OUTPUT
		retcode 	: UINT;
	END_VAR

  retcode := 0;

END_FUNCTION

#pragma warning (disable : 73)
FUNCTION VIRTUAL GLOBAL LseEasy::HmiScreenCreate
	VAR_INPUT
		screenno 	: UDINT;
	END_VAR

END_FUNCTION
#pragma warning (default : 73)

FUNCTION VIRTUAL GLOBAL LseEasy::EnglishFormatDateTime
	VAR_INPUT
		languageid 	: UDINT;
	END_VAR
	VAR_OUTPUT
		retcode 	: BOOL;
	END_VAR

  //  LOCAL_UNKNOWN             = 0x00,
  //  LOCAL_ARABIC              = 0x01,
  //  LOCAL_BULGARIAN           = 0x02,
  //  LOCAL_CATALAN             = 0x03,
  //  LOCAL_CHINESE             = 0x04,
  //  LOCAL_CZECH               = 0x05,
  //  LOCAL_DANISH              = 0x06,
  //  LOCAL_GERMAN              = 0x07,
  //  LOCAL_GREEK               = 0x08,
  //  LOCAL_ENGLISH             = 0x09,
  //  LOCAL_SPANISH             = 0x0A,
  //  LOCAL_FINNISH             = 0x0B,
  //  LOCAL_FRENCH              = 0x0C,
  //  LOCAL_HEBREW              = 0x0D,
  //  LOCAL_HUNGARIAN           = 0x0E,
  //  LOCAL_ICELANDIC           = 0x0F,
  //  LOCAL_ITALIAN             = 0x10,
  //  LOCAL_JAPANESE            = 0x11,
  //  LOCAL_KOREAN              = 0x12,
  //  LOCAL_DUTCH               = 0x13,
  //  LOCAL_NORWEGIAN           = 0x14,
  //  LOCAL_POLISH              = 0x15,
  //  LOCAL_PORTUGESE           = 0x16,
  //  LOCAL_ROMANIAN            = 0x18,
  //  LOCAL_RUSSIAN             = 0x19,
  //  LOCAL_CROATIA_SERBIAN     = 0x1A,
  //  LOCAL_SLOVAK              = 0x1B,
  //  LOCAL_ALBANIAN_MACEDONIAN = 0x1C,
  //  LOCAL_SWEDISH             = 0x1D,
  //  LOCAL_THAI                = 0x1E,
  //  LOCAL_TURKISH             = 0x1F,
  //  LOCAL_URDU                = 0x20,
  //  LOCAL_INDONESIAN          = 0x21,
  //  LOCAL_UKRAINIAN           = 0x22,
  //  LOCAL_BYELORUSSIAN        = 0x23,
  //  LOCAL_SLOVENIAN           = 0x24,
  //  LOCAL_ESTONIAN            = 0x25,
  //  LOCAL_LATVIAN             = 0x26,
  //  LOCAL_LITHUANIAN          = 0x27,
  //  LOCAL_FARSI               = 0x29,
  //  LOCAL_VIETNAMESE          = 0x2A,
  //  LOCAL_PASQUE              = 0x2D,
  //  LOCAL_AFRICAANS           = 0x36,
  //  LOCAL_GEORGIAN            = 0x37,
  //  LOCAL_FAEROESE            = 0x38,
  //  LOCAL_HINDI               = 0x39

  retcode := false;
  case(languageid and 16#FF) of
    16#00 : retcode := false; // unknown
//    16#09 : retcode := true; // english
  end_case;

END_FUNCTION

FUNCTION LseEasy::Create
	VAR_OUTPUT
		retcode 	: BOOL;
	END_VAR
  var
    anz  : udint;
    pline  : ^HMI_PRJINFO;
    dpne : array[0..80] of char;
  	pbox, fbox : ^void;
    pprj : ^_BOX_PROJECTLIST;
  end_var

  retcode := true; //false;

  // check actual selection of language
  if(HmiTextList.GetLanguageIndex(ActLanguage.Read()) = 16#FFFFFFFF) then
    ActLanguage.Write(0); // correct actual language
  end_if;

  HmiProject35.Start();

  HmiStateBit35.Start(this);
  HmiFunctionList35.Start();
  HmiShemeList35.Start(this);
  HmiVarList35.Start();
  HmiSetUpList35.Start();
  HmiTextList35.Start();
  HmiFont35.Start();
  HmiImage35.Start();
  HmiT9Config.Start();

  HmiProjectBegin(); // userinterface to add entries to div.list before lse-project is added

  // bootimage
  AddImageByIndex(HmiImageList.GetIndexByName(GetBootImage()), true);

  anz := HmiProjectList.GetNo();
  while(anz) do
    anz -= 1;
    pline := HmiProjectList.Get(anz);

    if(pline^.ima.ima = HMI_IMA_SCREEN) then
      MakePrjFileName(#dpne[0], #pline^.name[0]);
      if(HmiScreen.LoadFile(#dpne[0]) = true) then
        if(ScreenCreate(to_udint(pline^.ima.value)) = false) then
          retcode := false;
          OutMessageValue("ERROR: Create Screen ", to_udint(pline^.ima.value));
        end_if;
      else
        retcode := false;
        OutMessageValue("ERROR: Load Screen ", to_udint(pline^.ima.value));
      end_if;
    end_if;
    pline += sizeof(HMI_PRJINFO);
  end_while;

  HmiSetupList35.Create(CreateColor(HmiSetUpList.GetButColBack()),
                        CreateColor(HmiSetUpList.GetButColText()),
                        CreateColor(HmiSetUpList.GetTitleCol()),
                        CreateColor(HmiSetUpList.GetLimitCol()),
                        CreateColor(HmiSetUpList.GetWindowCol()),
                        CreateFrame(HmiSetUpList.GetButtonFrame(), 0),
                        CreateFrame(HmiSetUpList.GetWindowFrame(), 0),
                        UserProjectRevision(),
                        AddFont(HmiSetUpList.GetFontSchemeStandard()),
                        AddFont(HmiSetUpList.GetFontSchemeStandardSmall()));

  CreateAdd := true;
  HmiProjectCreate(); // userinterface to add entries to div.list
  CreateAdd := false;

  fbox := HmiFunctionList35.End(this); // functionlist als erstes machen weil ggf. Funktionsblöcke und Variablen noch addiert werden

  pbox := HmiVarList35.End();
  HmiProject35.AddEntry(BIGBOX_VARLIST, 0, pbox, false, false);

  pbox := HmiTextList35.End();
  HmiProject35.AddEntry(BIGBOX_TEXTLIST, 0, pbox, false, false);

  HmiProject35.AddEntry(BIGBOX_FUNCTIONLIST, 0, fbox, false, false);

  pbox := HmiShemeList35.End();
  HmiProject35.AddEntry(BIGBOX_SHEMELIST, 0, pbox, false, false);

  pbox := HmiSetupList35.End();
  HmiProject35.AddEntry(BIGBOX_SETUPLIST, 0, pbox, false, false);

  T9KeyboardConfig();
  pbox := HmiT9Config.End();
  if(pbox <> nil) then
    HmiProject35.AddEntry(BIGBOX_KEYBRD_T9, 0, pbox, false, false);
  end_if;

  if(HmiTextList35.GetErrorCnt() > 0) then
    OutMessage("ERROR: Maximum size of textlist reached");
    retcode := false;
  end_if;

  if(retcode = true) then

    ProjectBox := HmiProject35.End(HmiProjectList.GetStartScreen(), BackLightOff.Read(), TempInterval.Read());

    if(ProjectBox <> NIL) then
      pprj$^void := ProjectBox;
      HmiPrjCrc  := pprj^.boxhdr.crc32;

      // free furthermore unused memory
      HmiImageList.FreeMem();
      HmiFontList.FreeMem();
      // HmiTextList.FreeMem(); // xcomment: wunsch applikation 14.11.2017
      HmiFunctionList.FreeMem();
      HmiFontShemeList.FreeMem();
      HmiTextShemeList.FreeMem();
      HmiImageShemeList.FreeMem();
      HmiScreen.FreeMem();
    else
      retcode := false;
    end_if;
  end_if;

  if(retcode = false) then
    OutMessage("ERROR: Can't Create HMI-Project");
    SetErrorSvr(ErrCreateHmiProject);
  end_if;

//  SendProject(ProjectBox);
//  HmiProject35.Free();

END_FUNCTION

FUNCTION LseEasy::LoadProjectEntries
	VAR_OUTPUT
		retcode 	: BOOL;
	END_VAR
  var
    anz  : udint;
    pline  : ^HMI_PRJINFO;
    dpne : array[0..80] of char;
    state : bool;
  end_var

  retcode := true;
  anz     := HmiProjectList.GetNo();

  while(anz) do
    anz   -= 1;
    pline := HmiProjectList.Get(anz);
    state := true;

    case(pline^.ima.ima) of
      HMI_IMA_IMAGELIST      : MakePrjFileName(#dpne[0], #pline^.name[0]);
                               state := HmiImageList.LoadFile(#dpne[0]);
      HMI_IMA_SERVERLIST     : MakePrjFileName(#dpne[0], #pline^.name[0]);
                               state := HmiVarList.LoadFile(#dpne[0]);
                               HmiOverloadLight();
      HMI_IMA_FUNCTIONLIST   : MakePrjFileName(#dpne[0], #pline^.name[0]);
                               state := HmiFunctionList.LoadFile(#dpne[0]);
      HMI_IMA_GUIDEPOSTLIST  : MakePrjFileName(#dpne[0], #pline^.name[0]);
                               state := HmiTextList.LoadFile(#dpne[0], GetPrjPath(), ActLanguage.Read());
      HMI_IMA_TEXTSCHEMA     : MakePrjFileName(#dpne[0], #pline^.name[0]);
                               state := HmiTextShemeList.LoadFile(#dpne[0]);
      HMI_IMA_IMAGESCHEMA    : MakePrjFileName(#dpne[0], #pline^.name[0]);
                               state := HmiImageShemeList.LoadFile(#dpne[0]);
      HMI_IMA_FONTSCHEMA     : MakePrjFileName(#dpne[0], #pline^.name[0]);
                               state := HmiFontShemeList.LoadFile(#dpne[0]);
      HMI_IMA_UNITSCHEMA     : MakePrjFileName(#dpne[0], #pline^.name[0]);
                               state := HmiVarList.LoadUnitScheme(#dpne[0]);
      HMI_IMA_FONTLIST       : MakePrjFileName(#dpne[0], #pline^.name[0]);
                               state := HmiFontList.LoadFile(#dpne[0], GetPrjPath());
      HMI_IMA_COLORMAP       : MakePrjFileName(#dpne[0], #pline^.name[0]);
                               state := HmiColorMap.LoadFile(#dpne[0]);
      HMI_IMA_SETUPLIST      : MakePrjFileName(#dpne[0], #pline^.name[0]);
                               state := HmiSetUpList.LoadFile(#dpne[0]);
      HMI_IMA_CHKBITLIST     : MakePrjFileName(#dpne[0], #pline^.name[0]);
                               state := HmiChkBitList.LoadFile(#dpne[0]);

//      HMI_IMA_KEYPADLIST     : MakePrjFileName(#dpne[0], #pline^.name[0]);
//                           //GlobalKeypad.LoadFile(#dpne[0]);
    end_case;
    pline += sizeof(HMI_PRJINFO);

    if(state = false) then
      OutMessage("ERROR: Can't Load LSE-ProjectEntry");
      retcode := false;
      anz     := 0;
    end_if;

  end_while;

END_FUNCTION

FUNCTION LseEasy::LoadFile
	VAR_OUTPUT
		retcode 	: BOOL;
	END_VAR
  var
    dpne : array[0..80] of char;
    st : udint;
  end_var

  Free();

  retcode := false;

  MakePrjFileName(#dpne[0], HMI_PRJNAME);
  st := HmiProjectList.LoadFile(#dpne[0]);
  if(st = 1) then
    retcode := LoadProjectEntries();
  elsif(st = 2) then
    OutMessage("ERROR: Wrong LSE-Compiler Version");
    SetErrorSvr(ErrLseCompilerVersion);
  end_if;

  LseProjectRevision := HmiProjectList.GetLseProjectRevision();

  if(st <> 2) then
    if(retcode = false) then
      OutMessage("ERROR: Can't Load LSE-Project");
      SetErrorSvr(ErrLoadLseProject);
    end_if;
  end_if;

  if(retcode = true) then
    HmiVarList.SetLid(BacklightDimLid, HmiSwVersionLid, HmiHwVersionLid);
  end_if;

END_FUNCTION

FUNCTION LseEasy::ScreenCreate
	VAR_INPUT
		screennumber 	: UDINT;
	END_VAR
	VAR_OUTPUT
		retcode 	: BOOL;
	END_VAR
  VAR
  	anz, idx : udint;
    pany : ^HMI_ANYTHING;
    pctr : ^void;
    fct1, fct2 : uint;
  END_VAR

  fct1 := AddFunctionBlock(HmiScreen.GetStartFunct());
  fct2 := AddFunctionBlock(HmiScreen.GetEndFunct());

  ScreenStart(screennumber, fct1, fct2);

  anz := HmiScreen.GetZorderNo();
  idx := 0;
  while(anz) do
    pany := HmiScreen.GetZorder(idx);
    pctr := HmiScreen.GetControl(pany);

    if(pctr <> nil) then
      case pany^.ima of
        HMI_IMA_V_RECTANGLE : ScreenAddCtrlRectangle(pctr$^HMI_CTRL_RECTANGLE);
        HMI_IMA_V_LINE      : ScreenAddCtrlLine(pctr$^HMI_CTRL_LINE);
        HMI_IMA_V_CIRCLE    : ScreenAddCtrlCircle(pctr$^HMI_CTRL_CIRCLE);
        HMI_IMA_V_TEXT      : ScreenAddCtrlText(pctr$^HMI_CTRL_TEXT);
        HMI_IMA_V_IMAGE     : ScreenAddCtrlImage(pctr$^HMI_CTRL_IMAGE);
        HMI_IMA_V_IO        : ScreenAddCtrlIO(pctr$^HMI_CTRL_IO);
      end_case;
    end_if;

    anz -= 1;
    idx += 1;
  end_while;

  HmiScreenCreate(screennumber);

  retcode := ScreenStop(screennumber);

END_FUNCTION

FUNCTION LseEasy::GetFontInfo
	VAR_INPUT
		fontindex 	: UDINT;
	END_VAR
	VAR_OUTPUT
		retcode 	: ^HMI_FONTINFO;
	END_VAR
  VAR
  	pany : ^HMI_ANYTHING;
    lang : dint;
  END_VAR

  retcode := NIL;
  lang    := to_dint(HmiTextList.GetLanguageId(ActLanguage.Read()));
  pany    := HmiFontShemeList.GetResult(fontindex, lang);

  if(pany <> NIL) then
    if(pany^.ima = HMI_IMA_V_FONT) then
      retcode := HmiFontList.Get(pany^.value$udint);
    end_if;
  end_if;

END_FUNCTION

#define AttLEFT                   0x00 // horizontal alignment
#define AttCENTER                 0x10 // horizontal alignment
#define AttRIGHT                  0x20 // horizontal alignment
#define AttUP                     0x00 // vertical alignment
#define AttMID                    0x40 // vertical alignment
#define AttDOWN                   0x80 // vertical alignment
#define Att3D                     0x08 // used to display shade at each glyph
#define AttZOOM                   0x04 // zoom image
#define AttBOLD                   0x02 // used to display shade at each glyph

FUNCTION LseEasy::CreateAttrib
	VAR_INPUT
		att32 	: UDINT;
		fontindex 	: UDINT;
	END_VAR
	VAR_OUTPUT
		retcode 	: USINT;
	END_VAR
  VAR
    pfnt : ^HMI_FONTINFO;
  END_VAR

  retcode := 0;

  pfnt := GetFontInfo(fontindex);
  if(pfnt <> NIL) then
    if(pfnt^.attrib and T_STRIKEOUT) then
      retcode := retcode or ATT3D;
    end_if;
    if(pfnt^.attrib and T_BOLD) then
      retcode := retcode or AttBOLD;
    end_if;
  end_if;

  if(att32 and T_LEFTBOUND) then
    retcode := retcode or AttLEFT;
  end_if;
  if(att32 and T_CENTERBOUND) then
    retcode := retcode or AttCENTER;
  end_if;
  if(att32 and T_RIGHTBOUND) then
    retcode := retcode or AttRIGHT;
  end_if;
  if(att32 and T_UPBOUND) then
    retcode := retcode or AttUP;
  end_if;
  if(att32 and T_MIDBOUND) then
    retcode := retcode or AttMID;
  end_if;
  if(att32 and T_DOWNBOUND) then
    retcode := retcode or AttDOWN;
  end_if;

END_FUNCTION

FUNCTION LseEasy::CreateColor
	VAR_INPUT
		colindex 	: USINT;
	END_VAR
	VAR_OUTPUT
		retcode 	: UINT;
	END_VAR

  retcode := HmiColorMap.Get(colindex);

END_FUNCTION

FUNCTION LseEasy::CreateFrame
	VAR_INPUT
		frameindex 	: USINT;
		attrib 	: UDINT;
	END_VAR
	VAR_OUTPUT
		retcode 	: USINT;
	END_VAR

  retcode := frameindex;
  if(attrib and 16#20) then
    retcode := retcode or 16#80;
  end_if;

END_FUNCTION

FUNCTION LseEasy::CreateBarState
	VAR_INPUT
		attrib 	: UDINT;
	END_VAR
	VAR_OUTPUT
		retcode 	: USINT;
	END_VAR

  retcode := to_usint((attrib shr 24) and 7);
//    0 : // down->up
//    1 : // up->down
//    2 : // left->right
//    3 : // right->left
//    4 : // mid vertical
//    5 : // mid horizontal

END_FUNCTION
FUNCTION LseEasy::CreateMomStat
	VAR_INPUT
		pio 	: ^HMI_CTRL_IO;
	END_VAR
	VAR_OUTPUT
		retcode 	: UINT;
	END_VAR

  retcode := AddVariable(#pio^.server);
  if(retcode <> 16#FFFF) then
    if(pio^.act_momntry) then
      retcode := retcode or 16#8000;
    end_if;
  end_if;

END_FUNCTION

FUNCTION GLOBAL LseEasy::AddFunctionBlock
	VAR_INPUT
		functindex 	: UDINT;
	END_VAR
	VAR_OUTPUT
		retcode 	: UINT;
	END_VAR
  VAR
  	pfcb : ^HMI_FCTBLOCK;
  END_VAR

  retcode := 16#FFFF;

  pfcb$^void := HmiFunctionList.Get(functindex);
  if(pfcb <> NIL) then
    if(pfcb^.index35 <> HMI_DEFSCOPE) then
      retcode := pfcb^.index35$uint;
      return;
    end_if;

    retcode       := to_uint(HMIFunctionList35.AddEntry(pfcb));
    pfcb^.index35 := retcode;
  end_if;

END_FUNCTION

FUNCTION LseEasy::AddFunctionBlockIO
	VAR_INPUT
		pany 	: ^HMI_ANYTHING;
	END_VAR
	VAR_OUTPUT
		retcode 	: UINT;
	END_VAR

  retcode := 16#FFFF;
  if(pany^.ima = HMI_IMA_V_FUNCTIONLIST) then
    retcode := AddFunctionBlock(pany^.value$udint);
  end_if;

END_FUNCTION

FUNCTION LseEasy::AddVariable
	VAR_INPUT
		pany 	: ^HMI_ANYTHING;
	END_VAR
	VAR_OUTPUT
		retcode 	: UINT;
	END_VAR

  retcode := 16#FFFF;
  if(pany^.ima = HMI_IMA_V_SERVERLIST) then
    retcode := to_uint(HmiVarList.GetAdd35(pany^.value$udint));
  end_if;

END_FUNCTION

FUNCTION LseEasy::AddStateBitByName
	VAR_INPUT
		name 	: ^CHAR;
		invert 	: bool;
		access 	: UINT;
	END_VAR
	VAR_OUTPUT
		retcode 	: BOOL;
	END_VAR
  VAR
  	chkbit : HMI_CHKBIT;
    cno : udint;
    state : bool;
  END_VAR

  retcode := false;
  state   := (access <> 0);

  chkbit.no     := 16#FFFF;
  chkbit.invert := 0;

  cno := HmiChkBitList.GetChkBitIndex(name);
  if(cno < 16#FFFF) then
    chkbit.no := cno$uint;
    if(invert = true) then
      chkbit.invert := 1;
    end_if;
    state := true;
  end_if;

  if(state = true) then
    HmiStateBit35.AddEntry(#chkbit, access, NIL);
    retcode := true;
  end_if;

END_FUNCTION

FUNCTION LseEasy::AddVariableByName
  var_input
    name : ^char;
    station : udint;
  end_var
  var_output
    retcode : bool;
  end_var
  VAR
  	any : HMI_ANYTHING;
  END_VAR

  retcode := false;

  init_HMI_ANYTHING(#any);
  any.ima         := HMI_IMA_V_SERVERLIST;
  any.value$udint := HmiVarList.GetVarNoByName(name, station);
  if(AddVariable(#any) <> 16#FFFF) then
    retcode := true;
  end_if;

END_FUNCTION

FUNCTION LseEasy::GetLasalId
	VAR_INPUT
		pany 	: ^HMI_ANYTHING;
	END_VAR
	VAR_OUTPUT
		retcode 	: UDINT;
	END_VAR

  retcode := 0;
  if(pany^.ima = HMI_IMA_V_SERVERLIST) then
    retcode := HmiVarList.GetLasalId(pany^.value$udint);
  end_if;

END_FUNCTION

FUNCTION LseEasy::GetVariable
	VAR_INPUT
		pany 	: ^HMI_ANYTHING;
	END_VAR
	VAR_OUTPUT
		retcode 	: ^HMI_VARINFO;
	END_VAR

  retcode := nil;
  if(pany^.ima = HMI_IMA_V_SERVERLIST) then
    retcode := HmiVarList.Get(pany^.value$udint);
  end_if;

END_FUNCTION

FUNCTION LseEasy::AddSheme
	VAR_INPUT
		pany 	: ^HMI_ANYTHING;
	END_VAR
	VAR_OUTPUT
		retcode 	: UINT;
	END_VAR

  retcode := 16#FFFF;
  if(pany^.ima = HMI_IMA_V_IMAGESCHEMA) then
    retcode := HmiShemeList35.AddEntry(HmiImageShemeList.Get(to_udint(pany^.value)));
  elsif(pany^.ima = HMI_IMA_V_TEXTSCHEMA) then
    retcode := HmiShemeList35.AddEntry(HmiTextShemeList.Get(to_udint(pany^.value)));
  end_if;

END_FUNCTION

FUNCTION LseEasy::AddFont
	VAR_INPUT
		index 	: UDINT;
	END_VAR
	VAR_OUTPUT
		retcode 	: USINT;
	END_VAR
  VAR
    pfnt : ^HMI_FONTINFO;
    pbox : ^void;
  END_VAR

  retcode := 16#FF;

  pfnt := GetFontInfo(index);
  if(pfnt <> NIL) then
    if(pfnt^.index35 <> HMI_DEFSCOPE) then
      retcode := pfnt^.index35$usint;
      return;
    end_if;

    pbox := HmiFont35.CreateList(pfnt^.ptr, pfnt^.size);
    if(pbox <> NIL) then
      HmiFontList.SetIndex35(pfnt, HmiFontList.IncNumber());
      HmiProject35.AddEntry(BIGBOX_FONT, pfnt^.index35, pbox, false, true);
      retcode := pfnt^.index35$usint;
    end_if;
  end_if;

END_FUNCTION

FUNCTION LseEasy::AddText
	VAR_INPUT
		pany 	: ^HMI_ANYTHING;
	END_VAR
	VAR_OUTPUT
		retcode 	: UINT;
	END_VAR

  retcode := to_uint(HmiTextList.GetAdd35(pany));

END_FUNCTION

FUNCTION LseEasy::AddImageByIndex
	VAR_INPUT
		index 	: UDINT;
		bootimage 	: BOOL;
	END_VAR
	VAR_OUTPUT
		retcode 	: UINT;
	END_VAR
  VAR
  	pi : ^HMI_IMAGEINFO;
    pbox : ^void;
  END_VAR

  retcode := 16#FFFF;

  pi := HmiImageList.Get(index);
  if(pi <> NIL) then
    if(pi^.index35 <> HMI_DEFSCOPE) then
      retcode := pi^.index35$uint;
      return;
    end_if;

    pbox := HmiImage35.CreateList(pi^.width, pi^.height, pi^.transparent, pi^.state, pi^.datano, pi^.ptr);
    if(pbox <> NIL) then
      pi^.index35 := HmiImageList.IncNumber();
      if(bootimage = true) then
        HmiProject35.AddEntry(BIGBOX_BOOTIMAGE, pi^.index35, pbox, false, true);
      else
        HmiProject35.AddEntry(BIGBOX_IMAGE, pi^.index35, pbox, false, true);
      end_if;
      retcode := pi^.index35$uint;
    end_if;
  end_if;

END_FUNCTION

FUNCTION LseEasy::AddImage
	VAR_INPUT
		pany 	: ^HMI_ANYTHING;
	END_VAR
	VAR_OUTPUT
		retcode 	: UINT;
	END_VAR

  retcode := 16#FFFF;

  if(pany^.ima = HMI_IMA_V_IMAGELIST) then
    retcode := AddImageByIndex(pany^.value$udint, false);
  end_if;

END_FUNCTION

FUNCTION LseEasy::ScreenStart
	VAR_INPUT
		screennumber 	: UDINT;
		startfunct 	: UINT;
		endfunct 	: UINT;
	END_VAR

  StartScreen(to_uint(screennumber), startfunct, endfunct, CreateColor(HmiSetUpList.GetScreenColorBack()));

END_FUNCTION

FUNCTION LseEasy::ScreenAddCtrlRectangle
	VAR_INPUT
		ptr 	: ^HMI_CTRL_RECTANGLE;
	END_VAR
	VAR_OUTPUT
		retcode 	: BOOL;
	END_VAR
  VAR
  	sbit : usint;
  END_VAR

  retcode := false;

  sbit := HmiStateBit35.AddEntry(#ptr^.chkbit, 0, nil);
  if(AddScreen_CTRL_FRAME(ptr^.room.xy1.x, ptr^.room.xy1.y, ptr^.room.xy2.x, ptr^.room.xy2.y, CreateColor(ptr^.color), CreateFrame(ptr^.frame, ptr^.attrib), sbit) <> 0) then
    retcode := true;
  end_if;

END_FUNCTION

FUNCTION LseEasy::ScreenAddCtrlCircle
	VAR_INPUT
		ptr 	: ^HMI_CTRL_CIRCLE;
	END_VAR
	VAR_OUTPUT
		retcode 	: BOOL;
	END_VAR
  VAR
  	angle, arc : dint;
    xm, ym, rx, ry, r, a, ar : real;
    act, old : _XY;
    cdata : array[0..363] of _XY;
    cno : uint;
  	sbit : usint;
    pie : bool;
  END_VAR

  retcode := true;
  angle   := ptr^.angle / 10;
  arc     := ptr^.arc / 10;

  if(arc <> 0) then
    xm  := (to_real(ptr^.room.xy1.x + ptr^.room.xy2.x)) / 2;
    ym  := (to_real(ptr^.room.xy1.y + ptr^.room.xy2.y)) / 2;
    rx  := (to_real(ptr^.room.xy2.x - ptr^.room.xy1.x)) / 2;
    ry  := (to_real(ptr^.room.xy2.y - ptr^.room.xy1.y)) / 2;
    cno := 0;
    pie := true;

    if(arc >= 360) then
      arc := 360;
      pie := false;
    end_if;

    r := rx;
    if(ry > rx) then
      r  := ry;
    end_if;

    if(arc < 0) then
      angle += arc;
      arc   := -arc;
    end_if;

    a     := angle;
    old.x := -32768;
    old.y := -32768;
    arc   += 1;

    while(arc) do
      ar    := (a * 3.1416) / 180;
      act.x := to_int((COS(ar)    * rx) + xm + 0.5);
      act.y := to_int((-(SIN(ar)) * ry) + ym + 0.5);

      if((act.x <> old.x) | (act.y <> old.y)) then
        old := act;
        if(cno <= 360) then
          cdata[cno] := act;
          cno        += 1;
        end_if;
      end_if;

      a   += 1;
      arc -= 1;
    end_while;

    if(cno > 0) then
      if(pie = true) then
        cdata[cno].x := to_int(xm + 0.5);
        cdata[cno].y := to_int(ym + 0.5);
        cno += 1;
        cdata[cno] := cdata[0];
        cno += 1;
      end_if;

      sbit := HmiStateBit35.AddEntry(#ptr^.chkbit, 0, nil);
      if(AddScreen_CTRL_POLYLINE(#cdata[0], cno, CreateColor(ptr^.color), sbit) = 0) then
        retcode := false;
      end_if;
    end_if;
  end_if;

END_FUNCTION

FUNCTION LseEasy::ScreenAddCtrlLine
	VAR_INPUT
		ptr 	: ^HMI_CTRL_LINE;
	END_VAR
	VAR_OUTPUT
		retcode 	: BOOL;
	END_VAR
  VAR
  	sbit : usint;
  END_VAR

  retcode := false;
  sbit    := HmiStateBit35.AddEntry(#ptr^.chkbit, 0, nil);
  if(AddScreen_CTRL_POLYLINE(ptr^.ptxy$^_XY, ptr^.no, CreateColor(ptr^.color), sbit) <> 0) then
    retcode := true;
  end_if;

END_FUNCTION

FUNCTION LseEasy::ScreenAddCtrlImage
	VAR_INPUT
		ptr 	: ^HMI_CTRL_IMAGE;
	END_VAR
	VAR_OUTPUT
		retcode 	: BOOL;
	END_VAR
  VAR
  	sbit : usint;
  END_VAR

  retcode := false;
  sbit    := HmiStateBit35.AddEntry(#ptr^.chkbit, 0, nil);
  if(AddScreen_CTRL_IMAGE(ptr^.room.xy1.x, ptr^.room.xy1.y, ptr^.room.xy2.x, ptr^.room.xy2.y, AttMID or AttCENTER or AttZOOM, AddImage(#ptr^.any), sbit) <> 0) then
    retcode := true;
  end_if;

END_FUNCTION

FUNCTION LseEasy::ScreenAddCtrlText
	VAR_INPUT
		ptr 	: ^HMI_CTRL_TEXT;
	END_VAR
	VAR_OUTPUT
		retcode 	: BOOL;
	END_VAR
  VAR
  	txtidx : uint;
    sbit : usint;
  END_VAR

  retcode := false;

  if((ptr^.anything.ima = HMI_IMA_V_SERVERTEXT00) | (ptr^.anything.ima = HMI_IMA_V_SERVERUNITTEXT)) then
    if(HmiVarList.GetLasalId(ptr^.anything.value$udint) = 0) then
      return; // no valid lasalid --> do not add control
    end_if;
  end_if;

  sbit   := HmiStateBit35.AddEntry(#ptr^.chkbit, 0, #ptr^.anything);
  txtidx := AddText(#ptr^.anything);
  if(AddScreen_CTRL_TEXT(ptr^.room.xy1.x, ptr^.room.xy1.y, ptr^.room.xy2.x, ptr^.room.xy2.y,
                         CreateColor(ptr^.colorback), CreateColor(ptr^.colortext),
                         AddFont(ptr^.font), CreateAttrib(ptr^.attrib, ptr^.font),
                         CreateFrame(ptr^.frame, ptr^.attrib), txtidx, sbit) <> 0) then
    retcode := true;
  end_if;

END_FUNCTION

FUNCTION LseEasy::CreateVarConst
	VAR_INPUT
		vstate 	: ^USINT;
		pany 	: ^HMI_ANYTHING;
		pdata 	: ^HMI_ANYTHING;
		isog 	: BOOL;
		defval 	: DINT;
	END_VAR
	VAR_OUTPUT
		retcode 	: DINT;
	END_VAR
  VAR
  	varno : uint;
    pvar : ^HMI_VARINFO;
  END_VAR

  retcode := defval;
  vstate^ := 0;

  if(pany^.ima = HMI_IMA_V_SERVERLIST) then
    varno := AddVariable(pany);
    if(varno <> 0xFFFF) then
      retcode := varno;
      vstate^ := 1;
    end_if;
  elsif(pany^.ima = HMI_IMA_DINT_CONSTANT) then
    retcode := pany^.value;
  elsif(pdata <> NIL) then
    if(pdata^.ima = HMI_IMA_V_SERVERLIST) then
      pvar := HmiVarList.Get(pdata^.value$udint);
      if(pvar <> NIL) then
        pany := #pvar^.limit_lo;
        if(isog = true) then
          pany := #pvar^.limit_hi;
        end_if;
        retcode := CreateVarConst(vstate, pany, NIL, isog, defval);
      end_if;
    end_if;
  end_if;

END_FUNCTION

FUNCTION LseEasy::ScreenAddCtrlIO
	VAR_INPUT
		ptr 	: ^HMI_CTRL_IO;
	END_VAR
	VAR_OUTPUT
		retcode 	: BOOL;
	END_VAR
  VAR
  	st, lid  : udint;
    pvi : ^HMI_VARINFO;
    iot, dig, vugstate, vogstate, sbit : usint;
    vog, vug : dint;
    access, scmidx : uint;
  END_VAR

  retcode := false;
  st      := 1;

  access  := ptr^.access;
  if(ptr^.writeprotect = true) then
    access := 0;
  end_if;

  // todo: wenn access = 0 dann access von server holen

  case ptr^.iotype of
    HMI_IOT_NUMERIC:
      pvi := GetVariable(#ptr^.server);
      if(pvi <> nil) then

        lid  := GetLasalId(#ptr^.server);
        sbit := HmiStateBit35.AddEntry(#ptr^.chkbit, access, #ptr^.server);

        if((lid = TrendVal0Lid) | (lid = TrendVal1Lid)) then
          dig := 0;
          if(lid = TrendVal1Lid) then
            dig := 1;
          end_if;

          st := AddScreen_CTRL_OSZI(ptr^.room.xy1.x, ptr^.room.xy1.y, ptr^.room.xy2.x, ptr^.room.xy2.y,
                                    CreateColor(ptr^.color_back), CreateColor(ptr^.color_text),
                                    CreateAttrib(ptr^.attrib, ptr^.font),
                                    CreateFrame(ptr^.frame, ptr^.attrib),
                                    dig, sbit);
        elsif((lid = ListVal0Lid) | (lid = ListVal1Lid)) then
          dig := 0;
          if(lid = ListVal1Lid) then
            dig := 1;
          end_if;
          st := AddScreen_CTRL_LIST(ptr^.room.xy1.x, ptr^.room.xy1.y, ptr^.room.xy2.x, ptr^.room.xy2.y,
                                    AddVariable(#ptr^.server),
                                    CreateColor(ptr^.color_back), CreateColor(ptr^.color_text), CreateColor(9),
                                    AddFont(ptr^.font),
                                    CreateAttrib(ptr^.attrib, ptr^.font),
                                    CreateFrame(ptr^.frame, ptr^.attrib),
                                    dig, sbit);
        elsif(lid = PixMapLid) then
          st := AddScreen_CTRL_PIXMAP(ptr^.room.xy1.x, ptr^.room.xy1.y, ptr^.room.xy2.x, ptr^.room.xy2.y,
                                    CreateColor(ptr^.color_back), CreateColor(ptr^.color_text), 0, sbit);
        else

          case pvi^.vartype of
            HMI_DATE : iot := IOTYPE_DATE;
                       dig := DATEFORMAT_DDMMYYYY;
                       if(pvi^.subtype = 0) then
                         dig := DATEFORMAT_DDMM;
                       elsif(pvi^.subtype = 1) then
                         dig := DATEFORMAT_DDMMYY;
                       end_if;
                       if(EnglishFormatDateTime(HmiTextList.GetLanguageId(ActLanguage.Read())) = true) then
                         dig := dig or DATIM_USA;
                       end_if;
            HMI_TIME : iot := IOTYPE_TIME;
                       dig := TIMEFORMAT_HHMMSS;
                       if(pvi^.subtype = 0) then
                         dig := TIMEFORMAT_HHMM;
                       elsif(pvi^.subtype = 2) then
                         dig := TIMEFORMAT_MMSS;
                       end_if;
                       if(EnglishFormatDateTime(HmiTextList.GetLanguageId(ActLanguage.Read())) = true) then
                         dig := dig or DATIM_USA;
                       end_if;
            else       iot := IOTYPE_NUMERIC;
                       dig := HmiVarList.GetDigits(#ptr^.server, true);
          end_case;
